VAR_INPUT
  IN0 : INT ;
  IN1 : WORD ;
  IN2 : INT ;
  IN3 : INT ;
END_VAR
VAR_OUTPUT
  OUT4 : BOOL ;
  OUT5 : WORD ;
END_VAR
VAR
  STAT6 : STRUCT
   STAT7 : WORD ;
   STAT8 : WORD ;
   STAT9 : WORD ;
   STAT10 : BYTE ;
   STAT11 : BYTE ;
   STAT12 : BYTE ;
   STAT13 : BYTE ;
   STAT14 : BYTE ;
   STAT15 : BYTE ;
   STAT16 : BYTE ;
   STAT17 : BYTE ;
   STAT18 : BYTE ;
   STAT19 : BYTE ;
   STAT20 : BYTE ;
   STAT21 : BYTE ;
   STAT22 : BYTE ;
   STAT23 : BYTE ;
   STAT24 : BYTE ;
   STAT25 : BYTE ;
   STAT26 : BYTE ;
   STAT27 : BYTE ;
   STAT28 : BYTE ;
   STAT29 : BYTE ;
   STAT30 : BYTE ;
   STAT31 : BYTE ;
   STAT32 : BYTE ;
   STAT33 : BYTE ;
   STAT34 : BYTE ;
   STAT35 : BYTE ;
   STAT36 : BYTE ;
   STAT37 : BYTE ;
   STAT38 : BYTE ;
   STAT39 : BYTE ;
   STAT40 : BYTE ;
   STAT41 : BYTE ;
   STAT42 : BYTE ;
   STAT43 : BYTE ;
   STAT44 : BYTE ;
   STAT45 : BYTE ;
   STAT46 : BYTE ;
   STAT47 : BYTE ;
   STAT48 : BYTE ;
   STAT49 : BYTE ;
   STAT50 : BYTE ;
   STAT51 : BYTE ;
   STAT52 : BYTE ;
   STAT53 : BYTE ;
   STAT54 : BYTE ;
   STAT55 : BYTE ;
   STAT56 : BYTE ;
   STAT57 : BYTE ;
   STAT58 : BYTE ;
   STAT59 : BYTE ;
   STAT60 : BYTE ;
   STAT61 : BYTE ;
   STAT62 : BYTE ;
   STAT63 : BYTE ;
   STAT64 : BYTE ;
   STAT65 : BYTE ;
   STAT66 : BYTE ;
   STAT67 : BYTE ;
   STAT68 : BYTE ;
   STAT69 : BYTE ;
   STAT70 : BYTE ;
   STAT71 : BYTE ;
   STAT72 : BYTE ;
   STAT73 : BYTE ;
   STAT74 : BYTE ;
   STAT75 : BYTE ;
   STAT76 : BYTE ;
   STAT77 : BYTE ;
   STAT78 : BYTE ;
   STAT79 : BYTE ;
   STAT80 : BYTE ;
   STAT81 : BYTE ;
   STAT82 : BYTE ;
   STAT83 : BYTE ;
   STAT84 : BYTE ;
   STAT85 : BYTE ;
   STAT86 : BYTE ;
   STAT87 : BYTE ;
   STAT88 : BYTE ;
   STAT89 : BYTE ;
   STAT90 : BYTE ;
   STAT91 : BYTE ;
   STAT92 : BYTE ;
   STAT93 : BYTE ;
   STAT94 : BYTE ;
   STAT95 : BYTE ;
   STAT96 : BYTE ;
   STAT97 : BYTE ;
   STAT98 : BYTE ;
   STAT99 : BYTE ;
   STAT100 : BYTE ;
   STAT101 : BYTE ;
   STAT102 : BYTE ;
   STAT103 : BYTE ;
   STAT104 : BYTE ;
   STAT105 : BYTE ;
   STAT106 : BYTE ;
   STAT107 : BYTE ;
   STAT108 : BYTE ;
   STAT109 : BYTE ;
   STAT110 : BYTE ;
   STAT111 : BYTE ;
   STAT112 : BYTE ;
   STAT113 : BYTE ;
   STAT114 : BYTE ;
   STAT115 : BYTE ;
   STAT116 : BYTE ;
   STAT117 : BYTE ;
   STAT118 : BYTE ;
   STAT119 : BYTE ;
   STAT120 : BYTE ;
   STAT121 : BYTE ;
   STAT122 : BYTE ;
   STAT123 : BYTE ;
   STAT124 : BYTE ;
   STAT125 : BYTE ;
   STAT126 : BYTE ;
   STAT127 : BYTE ;
   STAT128 : BYTE ;
   STAT129 : BYTE ;
   STAT130 : BYTE ;
   STAT131 : BYTE ;
   STAT132 : BYTE ;
   STAT133 : BYTE ;
   STAT134 : BYTE ;
   STAT135 : BYTE ;
   STAT136 : BYTE ;
   STAT137 : BYTE ;
   STAT138 : BYTE ;
   STAT139 : BYTE ;
   STAT140 : BYTE ;
   STAT141 : BYTE ;
   STAT142 : BYTE ;
   STAT143 : BYTE ;
   STAT144 : BYTE ;
   STAT145 : BYTE ;
   STAT146 : BYTE ;
   STAT147 : BYTE ;
   STAT148 : BYTE ;
   STAT149 : BYTE ;
   STAT150 : BYTE ;
   STAT151 : BYTE ;
   STAT152 : BYTE ;
   STAT153 : BYTE ;
   STAT154 : BYTE ;
   STAT155 : BYTE ;
   STAT156 : BYTE ;
   STAT157 : BYTE ;
   STAT158 : BYTE ;
   STAT159 : BYTE ;
   STAT160 : BYTE ;
   STAT161 : BYTE ;
   STAT162 : BYTE ;
   STAT163 : BYTE ;
   STAT164 : BYTE ;
   STAT165 : BYTE ;
   STAT166 : BYTE ;
   STAT167 : BYTE ;
   STAT168 : BYTE ;
   STAT169 : BYTE ;
   STAT170 : BYTE ;
   STAT171 : BYTE ;
   STAT172 : BYTE ;
   STAT173 : BYTE ;
   STAT174 : BYTE ;
   STAT175 : BYTE ;
   STAT176 : BYTE ;
   STAT177 : BYTE ;
   STAT178 : BYTE ;
   STAT179 : BYTE ;
   STAT180 : BYTE ;
   STAT181 : BYTE ;
   STAT182 : BYTE ;
   STAT183 : BYTE ;
   STAT184 : BYTE ;
   STAT185 : BYTE ;
   STAT186 : BYTE ;
   STAT187 : BYTE ;
   STAT188 : BYTE ;
   STAT189 : BYTE ;
   STAT190 : BYTE ;
   STAT191 : BYTE ;
   STAT192 : BYTE ;
   STAT193 : BYTE ;
   STAT194 : BYTE ;
   STAT195 : BYTE ;
   STAT196 : BYTE ;
   STAT197 : BYTE ;
   STAT198 : BYTE ;
   STAT199 : BYTE ;
   STAT200 : BYTE ;
   STAT201 : BYTE ;
   STAT202 : BYTE ;
   STAT203 : BYTE ;
   STAT204 : BYTE ;
   STAT205 : BYTE ;
   STAT206 : BYTE ;
   STAT207 : BYTE ;
   STAT208 : BYTE ;
   STAT209 : BYTE ;
   STAT210 : BYTE ;
   STAT211 : BYTE ;
   STAT212 : BYTE ;
   STAT213 : BYTE ;
   STAT214 : BYTE ;
   STAT215 : BYTE ;
   STAT216 : BYTE ;
   STAT217 : BYTE ;
   STAT218 : BYTE ;
   STAT219 : BYTE ;
   STAT220 : BYTE ;
   STAT221 : BYTE ;
   STAT222 : BYTE ;
   STAT223 : BYTE ;
   STAT224 : BYTE ;
   STAT225 : BYTE ;
   STAT226 : BYTE ;
   STAT227 : BYTE ;
   STAT228 : BYTE ;
   STAT229 : BYTE ;
   STAT230 : BYTE ;
   STAT231 : BYTE ;
   STAT232 : BYTE ;
   STAT233 : BYTE ;
   STAT234 : BYTE ;
   STAT235 : BYTE ;
   STAT236 : BYTE ;
   STAT237 : BYTE ;
   STAT238 : BYTE ;
   STAT239 : BYTE ;
   STAT240 : BYTE ;
   STAT241 : BYTE ;
   STAT242 : BYTE ;
   STAT243 : BYTE ;
   STAT244 : BYTE ;
   STAT245 : BYTE ;
   STAT246 : BYTE ;
   STAT247 : BYTE ;
   STAT248 : BYTE ;
   STAT249 : BYTE ;
   STAT250 : BYTE ;
   STAT251 : BYTE ;
   STAT252 : BYTE ;
   STAT253 : BYTE ;
   STAT254 : BYTE ;
   STAT255 : BYTE ;
   STAT256 : BYTE ;
   STAT257 : BYTE ;
   STAT258 : BYTE ;
   STAT259 : BYTE ;
   STAT260 : BYTE ;
  END_STRUCT ;
  STAT261 : STRUCT
   STAT262 : WORD ;
   STAT263 : WORD ;
   STAT264 : WORD ;
   STAT265 : BYTE ;
   STAT266 : BYTE ;
   STAT267 : WORD ;
   STAT268 : WORD ;
   STAT269 : BYTE ;
   STAT270 : BYTE ;
   STAT271 : BYTE ;
   STAT272 : BYTE ;
   STAT273 : BYTE ;
   STAT274 : BYTE ;
   STAT275 : BYTE ;
   STAT276 : BYTE ;
   STAT277 : BYTE ;
   STAT278 : BYTE ;
   STAT279 : BYTE ;
   STAT280 : BYTE ;
   STAT281 : BYTE ;
   STAT282 : BYTE ;
   STAT283 : BYTE ;
   STAT284 : BYTE ;
   STAT285 : BYTE ;
   STAT286 : BYTE ;
   STAT287 : BYTE ;
   STAT288 : BYTE ;
   STAT289 : BYTE ;
   STAT290 : BYTE ;
   STAT291 : BYTE ;
   STAT292 : BYTE ;
   STAT293 : BYTE ;
   STAT294 : BYTE ;
   STAT295 : BYTE ;
   STAT296 : BYTE ;
   STAT297 : BYTE ;
   STAT298 : BYTE ;
   STAT299 : BYTE ;
   STAT300 : BYTE ;
   STAT301 : BYTE ;
   STAT302 : BYTE ;
   STAT303 : BYTE ;
   STAT304 : BYTE ;
   STAT305 : BYTE ;
   STAT306 : BYTE ;
   STAT307 : BYTE ;
   STAT308 : BYTE ;
   STAT309 : BYTE ;
   STAT310 : BYTE ;
   STAT311 : BYTE ;
   STAT312 : BYTE ;
   STAT313 : BYTE ;
   STAT314 : BYTE ;
   STAT315 : BYTE ;
   STAT316 : BYTE ;
   STAT317 : BYTE ;
   STAT318 : BYTE ;
   STAT319 : BYTE ;
   STAT320 : BYTE ;
   STAT321 : BYTE ;
   STAT322 : BYTE ;
   STAT323 : BYTE ;
   STAT324 : BYTE ;
   STAT325 : BYTE ;
   STAT326 : BYTE ;
   STAT327 : BYTE ;
   STAT328 : BYTE ;
   STAT329 : BYTE ;
   STAT330 : BYTE ;
   STAT331 : BYTE ;
   STAT332 : BYTE ;
   STAT333 : BYTE ;
   STAT334 : BYTE ;
   STAT335 : BYTE ;
   STAT336 : BYTE ;
   STAT337 : BYTE ;
   STAT338 : BYTE ;
   STAT339 : BYTE ;
   STAT340 : BYTE ;
   STAT341 : BYTE ;
   STAT342 : BYTE ;
   STAT343 : BYTE ;
   STAT344 : BYTE ;
   STAT345 : BYTE ;
   STAT346 : BYTE ;
   STAT347 : BYTE ;
   STAT348 : BYTE ;
   STAT349 : BYTE ;
   STAT350 : BYTE ;
   STAT351 : BYTE ;
   STAT352 : BYTE ;
   STAT353 : BYTE ;
   STAT354 : BYTE ;
   STAT355 : BYTE ;
   STAT356 : BYTE ;
   STAT357 : BYTE ;
   STAT358 : BYTE ;
   STAT359 : BYTE ;
   STAT360 : BYTE ;
   STAT361 : BYTE ;
   STAT362 : BYTE ;
   STAT363 : BYTE ;
   STAT364 : BYTE ;
   STAT365 : BYTE ;
   STAT366 : BYTE ;
   STAT367 : BYTE ;
   STAT368 : BYTE ;
   STAT369 : BYTE ;
   STAT370 : BYTE ;
   STAT371 : BYTE ;
   STAT372 : BYTE ;
   STAT373 : BYTE ;
   STAT374 : BYTE ;
   STAT375 : BYTE ;
   STAT376 : BYTE ;
   STAT377 : BYTE ;
   STAT378 : BYTE ;
   STAT379 : BYTE ;
   STAT380 : BYTE ;
   STAT381 : BYTE ;
   STAT382 : BYTE ;
   STAT383 : BYTE ;
   STAT384 : BYTE ;
   STAT385 : BYTE ;
   STAT386 : BYTE ;
   STAT387 : BYTE ;
   STAT388 : BYTE ;
   STAT389 : BYTE ;
   STAT390 : BYTE ;
   STAT391 : BYTE ;
   STAT392 : BYTE ;
   STAT393 : BYTE ;
   STAT394 : BYTE ;
   STAT395 : BYTE ;
   STAT396 : BYTE ;
   STAT397 : BYTE ;
   STAT398 : BYTE ;
   STAT399 : BYTE ;
   STAT400 : BYTE ;
   STAT401 : BYTE ;
   STAT402 : BYTE ;
   STAT403 : BYTE ;
   STAT404 : BYTE ;
   STAT405 : BYTE ;
   STAT406 : BYTE ;
   STAT407 : BYTE ;
   STAT408 : BYTE ;
   STAT409 : BYTE ;
   STAT410 : BYTE ;
   STAT411 : BYTE ;
   STAT412 : BYTE ;
   STAT413 : BYTE ;
   STAT414 : BYTE ;
   STAT415 : BYTE ;
   STAT416 : BYTE ;
   STAT417 : BYTE ;
   STAT418 : BYTE ;
   STAT419 : BYTE ;
   STAT420 : BYTE ;
   STAT421 : BYTE ;
   STAT422 : BYTE ;
   STAT423 : BYTE ;
   STAT424 : BYTE ;
   STAT425 : BYTE ;
   STAT426 : BYTE ;
   STAT427 : BYTE ;
   STAT428 : BYTE ;
   STAT429 : BYTE ;
   STAT430 : BYTE ;
   STAT431 : BYTE ;
   STAT432 : BYTE ;
   STAT433 : BYTE ;
   STAT434 : BYTE ;
   STAT435 : BYTE ;
   STAT436 : BYTE ;
   STAT437 : BYTE ;
   STAT438 : BYTE ;
   STAT439 : BYTE ;
   STAT440 : BYTE ;
   STAT441 : BYTE ;
   STAT442 : BYTE ;
   STAT443 : BYTE ;
   STAT444 : BYTE ;
   STAT445 : BYTE ;
   STAT446 : BYTE ;
   STAT447 : BYTE ;
   STAT448 : BYTE ;
   STAT449 : BYTE ;
   STAT450 : BYTE ;
   STAT451 : BYTE ;
   STAT452 : BYTE ;
   STAT453 : BYTE ;
   STAT454 : BYTE ;
   STAT455 : BYTE ;
   STAT456 : BYTE ;
   STAT457 : BYTE ;
   STAT458 : BYTE ;
   STAT459 : BYTE ;
   STAT460 : BYTE ;
   STAT461 : BYTE ;
   STAT462 : BYTE ;
   STAT463 : BYTE ;
   STAT464 : BYTE ;
   STAT465 : BYTE ;
   STAT466 : BYTE ;
   STAT467 : BYTE ;
   STAT468 : BYTE ;
   STAT469 : BYTE ;
   STAT470 : BYTE ;
   STAT471 : BYTE ;
   STAT472 : BYTE ;
   STAT473 : BYTE ;
   STAT474 : BYTE ;
   STAT475 : BYTE ;
   STAT476 : BYTE ;
   STAT477 : BYTE ;
   STAT478 : BYTE ;
   STAT479 : BYTE ;
   STAT480 : BYTE ;
   STAT481 : BYTE ;
   STAT482 : BYTE ;
   STAT483 : BYTE ;
   STAT484 : BYTE ;
   STAT485 : BYTE ;
   STAT486 : BYTE ;
   STAT487 : BYTE ;
   STAT488 : BYTE ;
   STAT489 : BYTE ;
   STAT490 : BYTE ;
   STAT491 : BYTE ;
   STAT492 : BYTE ;
   STAT493 : BYTE ;
   STAT494 : BYTE ;
   STAT495 : BYTE ;
   STAT496 : BYTE ;
   STAT497 : BYTE ;
   STAT498 : BYTE ;
   STAT499 : BYTE ;
   STAT500 : BYTE ;
   STAT501 : BYTE ;
   STAT502 : BYTE ;
   STAT503 : BYTE ;
   STAT504 : BYTE ;
   STAT505 : BYTE ;
   STAT506 : BYTE ;
   STAT507 : BYTE ;
   STAT508 : BYTE ;
   STAT509 : BYTE ;
   STAT510 : BYTE ;
   STAT511 : BYTE ;
   STAT512 : BYTE ;
   STAT513 : BYTE ;
   STAT514 : BYTE ;
  END_STRUCT ;
  STAT515 : INT ;
  STAT516 : INT ;
  STAT517 : BOOL ;
  STAT518 : BOOL ;
  STAT519 : BOOL ;
  STAT520 : BOOL ;
  STAT521 : WORD ;
  STAT522 : INT ;
  STAT523 : BOOL ;
  STAT524 : BOOL ;
  STAT525 : WORD ;
  STAT526 : INT ;
  STAT527 : INT ;
  STAT528 : BOOL ;
  STAT529 : BOOL ;
  STAT530 : WORD ;
  STAT531 : BOOL ;
  STAT532 : WORD ;
  STAT533 : "TON";
  STAT541 : BOOL ;
  STAT542 : BOOL ;
  STAT543 : BOOL ;
  STAT544 : WORD ;
END_VAR
VAR_TEMP
  TEMP545 : ANY ;
  TEMP546 : ANY ;
  TEMP547 : INT ;
  TEMP548 : DWORD ;
  TEMP549 : DWORD ;
END_VAR
BEGIN
NETWORK
TITLE =
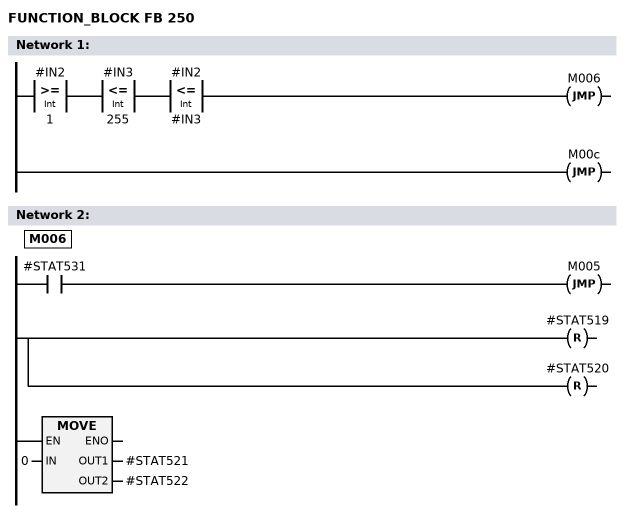

      SET   ;
      A(    ;
      L     #IN2;
      L     1;
      >=I   ;
      )     ;
      A(    ;
      L     #IN3;
      L     255;
      <=I   ;
      )     ;
      A(    ;
      L     #IN2;
      L     #IN3;
      <=I   ;
      )     ;
      JC    M006;
      JU    M00c;
NETWORK
TITLE =

M006: A     #STAT531;
      JC    M005;
      SET   ;
      R     #STAT519;
      R     #STAT520;
      L     0;
      T     #STAT521;
      T     #STAT522;
NETWORK
TITLE =

      LAR1  P##TEMP545;
      L     B#16#10;
      T     LB [AR1,P#0.0];
      L     B#16#2;
      T     LB [AR1,P#1.0];
      L     6;
      T     LW [AR1,P#2.0];
      L     DINO;
      T     LW [AR1,P#4.0];
      L     270;
      L     8;
      *I    ;
      L     P#DBX 0.0;
      +D    ;
      T     LD [AR1,P#6.0];
NETWORK
TITLE =
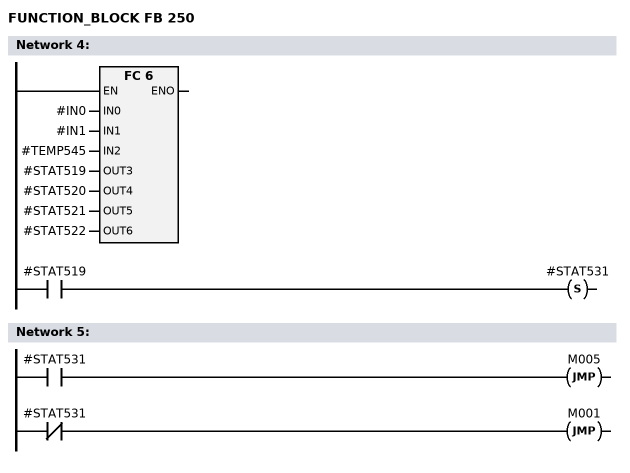

      CALL FC     6 (
           IN0                      := #IN0,
           IN1                      := #IN1,
           IN2                      := #TEMP545,
           OUT3                     := #STAT519,
           OUT4                     := #STAT520,
           OUT5                     := #STAT521,
           OUT6                     := #STAT522);
      SET   ;
      A     #STAT519;
      S     #STAT531;
NETWORK
TITLE =

      A     #STAT531;
      JC    M005;
      AN    #STAT531;
      JC    M001;
NETWORK
TITLE =

M005: LAR1  P##TEMP546;
      L     B#16#10;
      T     LB [AR1,P#0.0];
      L     B#16#2;
      T     LB [AR1,P#1.0];
      L     DIW  274;
      T     LW [AR1,P#2.0];
      L     DINO;
      T     LW [AR1,P#4.0];
      L     276;
      L     8;
      *I    ;
      L     P#DBX 0.0;
      +D    ;
      T     LD [AR1,P#6.0];
NETWORK
TITLE =
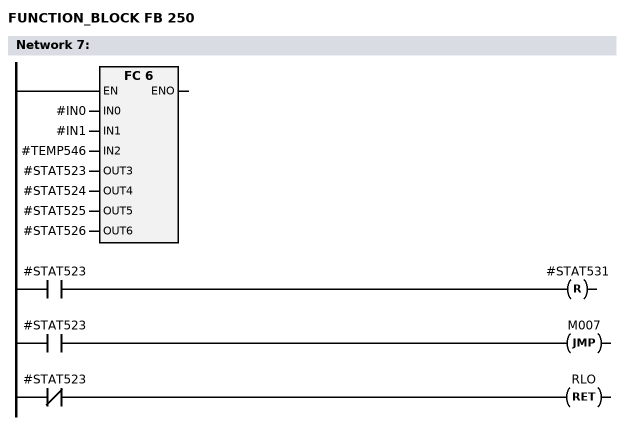

      CALL FC     6 (
           IN0                      := #IN0,
           IN1                      := #IN1,
           IN2                      := #TEMP546,
           OUT3                     := #STAT523,
           OUT4                     := #STAT524,
           OUT5                     := #STAT525,
           OUT6                     := #STAT526);
      SET   ;
      A     #STAT523;
      R     #STAT531;
      A     #STAT523;
      JC    M007;
      AN    #STAT523;
      BEC   ;
NETWORK
TITLE =

M007: SET   ;
      L     #STAT261.STAT266;
      L     3;
      ==I   ;
      =     #STAT517;
      L     #STAT261.STAT266;
      L     16;
      ==I   ;
      =     #STAT518;
      A     #STAT517;
      JC    M00b;
      A     #STAT518;
      JC    M009;
      JU    M008;
NETWORK
TITLE =

M00b: O(    ;
      L     #STAT261.STAT268;
      L     1;
      <I    ;
      )     ;
      O(    ;
      L     #STAT261.STAT268;
      L     100;
      >I    ;
      )     ;
      JC    M00a;
      L     #STAT261.STAT267;
      SRW   8;
      T     #TEMP547;
      L     #IN2;
      L     #TEMP547;
      +I    ;
      T     #TEMP547;
      O(    ;
      L     #TEMP547;
      L     #IN2;
      <I    ;
      )     ;
      O(    ;
      L     #TEMP547;
      L     #IN3;
      >I    ;
      )     ;
      JC    M00a;
      L     #STAT261.STAT262;
      T     #STAT6.STAT7;
      L     #STAT261.STAT263;
      T     #STAT6.STAT8;
      L     #STAT261.STAT265;
      T     #STAT6.STAT10;
      L     #STAT261.STAT266;
      T     #STAT6.STAT11;
      L     #STAT261.STAT268;
      SLW   1;
      T     #STAT6.STAT12;
      L     #STAT6.STAT12;
      +     3;
      T     #STAT6.STAT9;
      OPN   DB [#TEMP547];
      L     #STAT261.STAT267;
      SLW   8;
      SRW   8;
      SLD   4;
      T     #TEMP548;
      L     P##STAT6;
      L     P#9.0;
      +D    ;
      T     #TEMP549;
      L     #STAT261.STAT268;
M003: T     #STAT532;
      L     DBW [#TEMP548];
      T     DIW [#TEMP549];
      L     #TEMP548;
      +     16;
      T     #TEMP548;
      L     #TEMP549;
      +     16;
      T     #TEMP549;
      L     #STAT532;
      LOOP  M003;
      L     #STAT6.STAT9;
      +     6;
      T     #STAT527;
      L     W#16#0;
      T     #OUT5;
      R     #OUT4;
      S     #STAT543;
      JU    M001;
NETWORK
TITLE =

M009: O(    ;
      L     #STAT261.STAT268;
      L     1;
      <I    ;
      )     ;
      O(    ;
      L     #STAT261.STAT268;
      L     100;
      >I    ;
      )     ;
      JC    M00a;
      L     #STAT261.STAT267;
      T     #STAT6.STAT15;
      SRW   8;
      T     #STAT6.STAT12;
      T     #TEMP547;
      L     #IN2;
      L     #TEMP547;
      +I    ;
      T     #TEMP547;
      O(    ;
      L     #TEMP547;
      L     #IN2;
      <I    ;
      )     ;
      O(    ;
      L     #TEMP547;
      L     #IN3;
      >I    ;
      )     ;
      JC    M00a;
      L     #STAT261.STAT262;
      T     #STAT6.STAT7;
      L     #STAT261.STAT263;
      T     #STAT6.STAT8;
      L     #STAT261.STAT265;
      T     #STAT6.STAT10;
      L     #STAT261.STAT266;
      T     #STAT6.STAT11;
      L     6;
      T     #STAT6.STAT9;
      L     0;
      T     #STAT6.STAT14;
      L     #STAT261.STAT268;
      T     #STAT6.STAT15;
      OPN   DB [#TEMP547];
      L     #STAT261.STAT267;
      SLW   8;
      SRW   8;
      T     #STAT6.STAT13;
      SLD   4;
      T     #TEMP549;
      L     P##STAT261;
      L     P#13.0;
      +D    ;
      T     #TEMP548;
      L     #STAT261.STAT268;
M004: T     #STAT532;
      L     DIW [#TEMP548];
      T     DBW [#TEMP549];
      L     #TEMP548;
      +     16;
      T     #TEMP548;
      L     #TEMP549;
      +     16;
      T     #TEMP549;
      L     #STAT532;
      LOOP  M004;
      L     12;
      T     #STAT527;
      L     W#16#0;
      T     #OUT5;
      R     #OUT4;
      S     #STAT543;
      JU    M001;
NETWORK
TITLE =

M00c: L     W#16#290;
      T     #OUT5;
      S     #OUT4;
      BEU   ;
M008: L     B#16#1;
      T     #STAT6.STAT12;
      L     W#16#300;
      T     #OUT5;
      JU    M002;
M00a: L     B#16#2;
      T     #STAT6.STAT12;
      L     W#16#381;
      T     #OUT5;
      JU    M002;
M002: L     #STAT261.STAT262;
      T     #STAT6.STAT7;
      L     #STAT261.STAT263;
      T     #STAT6.STAT8;
      L     #STAT261.STAT265;
      T     #STAT6.STAT10;
      L     #STAT261.STAT266;
      +     B#16#80;
      T     #STAT6.STAT11;
      L     3;
      T     #STAT6.STAT9;
      L     9;
      T     #STAT527;
      S     #OUT4;
      S     #STAT543;
      JU    M001;
NETWORK
TITLE =

M001: CALL FC     5 (
           IN0                      := #STAT543,
           IN1                      := #IN0,
           IN2                      := #IN1,
           IN3                      := #STAT6,
           IN4                      := #STAT527,
           OUT5                     := #STAT528,
           OUT6                     := #STAT529,
           OUT7                     := #STAT530);
      SET   ;
      R     #STAT543;
      BEU   ;
END_FUNCTION_BLOCK

FUNCTION FC 14 : VOID
VERSION : 0.1

BEGIN
NETWORK
TITLE =

      CALL FB   250 , DB   250 (
           IN0                      := 1,
           IN1                      := W#16#180,
           IN2                      := 95,
           IN3                      := 95,
           OUT4                     := DB250.DBX    8.0,
           OUT5                     := DB250.DBW   10);
      NOP   0;
NETWORK
TITLE =

      A     I      0.0;
      =     DB95.DBX    1.0;
NETWORK
TITLE =

      A     Q    160.6;
      =     DB95.DBX    1.1;
NETWORK
TITLE =

      A(    ;
      L     DB51.DBD  252;
      L     1.000000e+003;
      *R    ;
      T     MD   100;
      AN    OV;
      SAVE  ;
      CLR   ;
      A     BR;
      )     ;
      JNB   M001;
      L     MD   100;
      RND   ;
      T     DB95.DBW   18;
M001: NOP   0;
NETWORK
TITLE =

      A(    ;
      L     DB51.DBD  292;
      L     1.000000e+003;
      *R    ;
      T     MD   104;
      AN    OV;
      SAVE  ;
      CLR   ;
      A     BR;
      )     ;
      JNB   M002;
      L     MD   104;
      RND   ;
      T     DB95.DBW   20;
M002: NOP   0;
NETWORK
TITLE =

      A(    ;
      L     DB51.DBD   92;
      L     1.000000e+003;
      *R    ;
      T     MD   108;
      AN    OV;
      SAVE  ;
      CLR   ;
      A     BR;
      )     ;
      JNB   M003;
      L     MD   108;
      RND   ;
      T     DB95.DBW   22;
M003: NOP   0;
NETWORK
TITLE =

      A(    ;
      L     DB51.DBD  212;
      L     1.000000e+003;
      *R    ;
      T     MD   112;
      AN    OV;
      SAVE  ;
      CLR   ;
      A     BR;
      )     ;
      JNB   M004;
      L     MD   112;
      RND   ;
      T     DB95.DBW   24;
M004: NOP   0;
NETWORK
TITLE =

      A(    ;
      L     DB51.DBD   52;
      L     1.000000e+003;
      *R    ;
      T     MD   116;
      AN    OV;
      SAVE  ;
      CLR   ;
      A     BR;
      )     ;
      JNB   M005;
      L     MD   116;
      RND   ;
      T     DB95.DBW   26;
M005: NOP   0;
NETWORK
TITLE =

      A(    ;
      L     DB51.DBD  172;
      L     1.000000e+003;
      *R    ;
      T     MD   120;
      AN    OV;
      SAVE  ;
      CLR   ;
      A     BR;
      )     ;
      JNB   M006;
      L     MD   120;
      RND   ;
      T     DB95.DBW   28;
M006: NOP   0;
NETWORK
TITLE =

      A(    ;
      L     DB51.DBD   12;
      L     1.000000e+003;
      *R    ;
      T     MD   124;
      AN    OV;
      SAVE  ;
      CLR   ;
      A     BR;
      )     ;
      JNB   M007;
      L     MD   124;
      RND   ;
      T     DB95.DBW   30;
M007: NOP   0;
NETWORK
TITLE =

      A(    ;
      L     DB51.DBD  132;
      L     1.000000e+003;
      *R    ;
      T     MD   128;
      AN    OV;
      SAVE  ;
      CLR   ;
      A     BR;
      )     ;
      JNB   M008;
      L     MD   128;
      RND   ;
      T     DB95.DBW   32;
M008: NOP   0;
NETWORK
TITLE =

      A(    ;
      L     DB51.DBD  256;
      L     1.000000e+003;
      *R    ;
      T     MD   132;
      AN    OV;
      SAVE  ;
      CLR   ;
      A     BR;
      )     ;
      JNB   M009;
      L     MD   132;
      RND   ;
      T     DB95.DBW   38;
M009: NOP   0;
NETWORK
TITLE =

      A(    ;
      L     DB51.DBD  296;
      L     1.000000e+003;
      *R    ;
      T     MD   136;
      AN    OV;
      SAVE  ;
      CLR   ;
      A     BR;
      )     ;
      JNB   M00a;
      L     MD   136;
      RND   ;
      T     DB95.DBW   40;
M00a: NOP   0;
NETWORK
TITLE =

      A(    ;
      L     DB51.DBD   96;
      L     1.000000e+003;
      *R    ;
      T     MD   140;
      AN    OV;
      SAVE  ;
      CLR   ;
      A     BR;
      )     ;
      JNB   M00b;
      L     MD   140;
      RND   ;
      T     DB95.DBW   42;
M00b: NOP   0;
NETWORK
TITLE =

      A(    ;
      L     DB51.DBD  216;
      L     1.000000e+003;
      *R    ;
      T     MD   144;
      AN    OV;
      SAVE  ;
      CLR   ;
      A     BR;
      )     ;
      JNB   M00c;
      L     MD   144;
      RND   ;
      T     DB95.DBW   44;
M00c: NOP   0;
NETWORK
TITLE =

      A(    ;
      L     DB51.DBD   56;
      L     1.000000e+003;
      *R    ;
      T     MD   148;
      AN    OV;
      SAVE  ;
      CLR   ;
      A     BR;
      )     ;
      JNB   M00d;
      L     MD   148;
      RND   ;
      T     DB95.DBW   46;
M00d: NOP   0;
NETWORK
TITLE =

      A(    ;
      L     DB51.DBD  176;
      L     1.000000e+003;
      *R    ;
      T     MD   152;
      AN    OV;
      SAVE  ;
      CLR   ;
      A     BR;
      )     ;
      JNB   M00e;
      L     MD   152;
      RND   ;
      T     DB95.DBW   48;
M00e: NOP   0;
NETWORK
TITLE =

      A(    ;
      L     DB51.DBD   16;
      L     1.000000e+003;
      *R    ;
      T     MD   156;
      AN    OV;
      SAVE  ;
      CLR   ;
      A     BR;
      )     ;
      JNB   M00f;
      L     MD   156;
      RND   ;
      T     DB95.DBW   50;
M00f: NOP   0;
NETWORK
TITLE =

      A(    ;
      L     DB51.DBD  136;
      L     1.000000e+003;
      *R    ;
      T     MD   160;
      AN    OV;
      SAVE  ;
      CLR   ;
      A     BR;
      )     ;
      JNB   M010;
      L     MD   160;
      RND   ;
      T     DB95.DBW   52;
M010: NOP   0;
NETWORK
TITLE =

      A(    ;
      L     DB51.DBD  260;
      L     1.000000e+003;
      *R    ;
      T     MD   164;
      AN    OV;
      SAVE  ;
      CLR   ;
      A     BR;
      )     ;
      JNB   M011;
      L     MD   164;
      RND   ;
      T     DB95.DBW   58;
M011: NOP   0;
NETWORK
TITLE =

      A(    ;
      L     DB51.DBD  300;
      L     1.000000e+003;
      *R    ;
      T     MD   168;
      AN    OV;
      SAVE  ;
      CLR   ;
      A     BR;
      )     ;
      JNB   M012;
      L     MD   168;
      RND   ;
      T     DB95.DBW   60;
M012: NOP   0;
NETWORK
TITLE =

      A(    ;
      L     DB51.DBD  100;
      L     1.000000e+003;
      *R    ;
      T     MD   172;
      AN    OV;
      SAVE  ;
      CLR   ;
      A     BR;
      )     ;
      JNB   M013;
      L     MD   172;
      RND   ;
      T     DB95.DBW   62;
M013: NOP   0;
NETWORK
TITLE =

      A(    ;
      L     DB51.DBD  220;
      L     1.000000e+003;
      *R    ;
      T     MD   176;
      AN    OV;
      SAVE  ;
      CLR   ;
      A     BR;
      )     ;
      JNB   M014;
      L     MD   176;
      RND   ;
      T     DB95.DBW   64;
M014: NOP   0;
NETWORK
TITLE =

      A(    ;
      L     DB51.DBD   60;
      L     1.000000e+003;
      *R    ;
      T     MD   180;
      AN    OV;
      SAVE  ;
      CLR   ;
      A     BR;
      )     ;
      JNB   M015;
      L     MD   180;
      RND   ;
      T     DB95.DBW   66;
M015: NOP   0;
NETWORK
TITLE =

      A(    ;
      L     DB51.DBD  180;
      L     1.000000e+003;
      *R    ;
      T     MD   184;
      AN    OV;
      SAVE  ;
      CLR   ;
      A     BR;
      )     ;
      JNB   M016;
      L     MD   184;
      RND   ;
      T     DB95.DBW   68;
M016: NOP   0;
NETWORK
TITLE =

      A(    ;
      L     DB51.DBD   20;
      L     1.000000e+003;
      *R    ;
      T     MD   188;
      AN    OV;
      SAVE  ;
      CLR   ;
      A     BR;
      )     ;
      JNB   M017;
      L     MD   188;
      RND   ;
      T     DB95.DBW   70;
M017: NOP   0;
NETWORK
TITLE =

      A(    ;
      L     DB51.DBD  140;
      L     1.000000e+003;
      *R    ;
      T     MD   192;
      AN    OV;
      SAVE  ;
      CLR   ;
      A     BR;
      )     ;
      JNB   M018;
      L     MD   192;
      RND   ;
      T     DB95.DBW   72;
M018: NOP   0;
NETWORK
TITLE =

      A(    ;
      L     DB51.DBD  264;
      L     1.000000e+003;
      *R    ;
      T     MD   296;
      AN    OV;
      SAVE  ;
      CLR   ;
      A     BR;
      )     ;
      JNB   M019;
      L     MD   296;
      RND   ;
      T     DB95.DBW   78;
M019: NOP   0;
NETWORK
TITLE =

      A(    ;
      L     DB51.DBD  304;
      L     1.000000e+003;
      *R    ;
      T     MD   304;
      AN    OV;
      SAVE  ;
      CLR   ;
      A     BR;
      )     ;
      JNB   M01a;
      L     MD   304;
      RND   ;
      T     DB95.DBW   80;
M01a: NOP   0;
NETWORK
TITLE =

      A(    ;
      L     DB51.DBD  104;
      L     1.000000e+003;
      *R    ;
      T     MD   308;
      AN    OV;
      SAVE  ;
      CLR   ;
      A     BR;
      )     ;
      JNB   M01b;
      L     MD   308;
      RND   ;
      T     DB95.DBW   82;
M01b: NOP   0;
NETWORK
TITLE =

      A(    ;
      L     DB51.DBD  224;
      L     1.000000e+003;
      *R    ;
      T     MD   312;
      AN    OV;
      SAVE  ;
      CLR   ;
      A     BR;
      )     ;
      JNB   M01c;
      L     MD   312;
      RND   ;
      T     DB95.DBW   84;
M01c: NOP   0;
NETWORK
TITLE =

      A(    ;
      L     DB51.DBD   64;
      L     1.000000e+003;
      *R    ;
      T     MD   316;
      AN    OV;
      SAVE  ;
      CLR   ;
      A     BR;
      )     ;
      JNB   M01d;
      L     MD   316;
      RND   ;
      T     DB95.DBW   86;
M01d: NOP   0;
NETWORK
TITLE =

      A(    ;
      L     DB51.DBD  184;
      L     1.000000e+003;
      *R    ;
      T     MD   320;
      AN    OV;
      SAVE  ;
      CLR   ;
      A     BR;
      )     ;
      JNB   M01e;
      L     MD   320;
      RND   ;
      T     DB95.DBW   88;
M01e: NOP   0;
NETWORK
TITLE =

      A(    ;
      L     DB51.DBD   24;
      L     1.000000e+003;
      *R    ;
      T     MD   324;
      AN    OV;
      SAVE  ;
      CLR   ;
      A     BR;
      )     ;
      JNB   M01f;
      L     MD   324;
      RND   ;
      T     DB95.DBW   90;
M01f: NOP   0;
NETWORK
TITLE =

      A(    ;
      L     DB51.DBD  144;
      L     1.000000e+003;
      *R    ;
      T     MD   328;
      AN    OV;
      SAVE  ;
      CLR   ;
      A     BR;
      )     ;
      JNB   M020;
      L     MD   328;
      RND   ;
      T     DB95.DBW   92;
M020: NOP   0;
END_FUNCTION

FUNCTION FC 1 : VOID
VERSION : 0.1

BEGIN
NETWORK
TITLE =
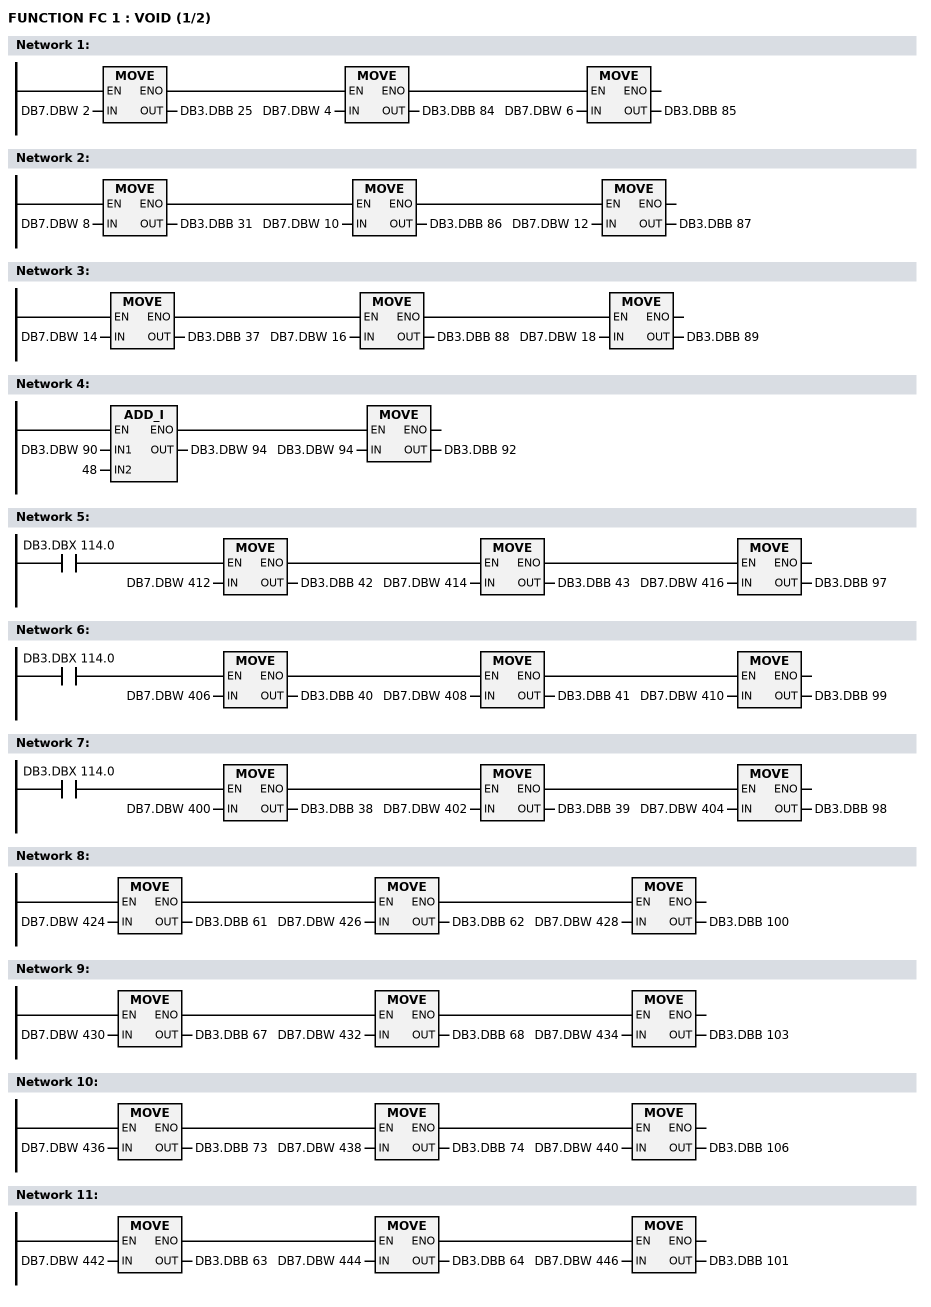

      A(    ;
      A(    ;
      L     DB7.DBW    2;
      T     DB3.DBB   25;
      SET   ;
      SAVE  ;
      CLR   ;
      A     BR;
      )     ;
      JNB   M001;
      L     DB7.DBW    4;
      T     DB3.DBB   84;
      SET   ;
      SAVE  ;
      CLR   ;
M001: A     BR;
      )     ;
      JNB   M002;
      L     DB7.DBW    6;
      T     DB3.DBB   85;
M002: NOP   0;
NETWORK
TITLE =

      A(    ;
      A(    ;
      L     DB7.DBW    8;
      T     DB3.DBB   31;
      SET   ;
      SAVE  ;
      CLR   ;
      A     BR;
      )     ;
      JNB   M003;
      L     DB7.DBW   10;
      T     DB3.DBB   86;
      SET   ;
      SAVE  ;
      CLR   ;
M003: A     BR;
      )     ;
      JNB   M004;
      L     DB7.DBW   12;
      T     DB3.DBB   87;
M004: NOP   0;
NETWORK
TITLE =

      A(    ;
      A(    ;
      L     DB7.DBW   14;
      T     DB3.DBB   37;
      SET   ;
      SAVE  ;
      CLR   ;
      A     BR;
      )     ;
      JNB   M005;
      L     DB7.DBW   16;
      T     DB3.DBB   88;
      SET   ;
      SAVE  ;
      CLR   ;
M005: A     BR;
      )     ;
      JNB   M006;
      L     DB7.DBW   18;
      T     DB3.DBB   89;
M006: NOP   0;
NETWORK
TITLE =

      A(    ;
      L     DB3.DBW   90;
      L     48;
      +I    ;
      T     DB3.DBW   94;
      AN    OV;
      SAVE  ;
      CLR   ;
      A     BR;
      )     ;
      JNB   M007;
      L     DB3.DBW   94;
      T     DB3.DBB   92;
M007: NOP   0;
NETWORK
TITLE =

      A(    ;
      A(    ;
      A     DB3.DBX  114.0;
      JNB   M008;
      L     DB7.DBW  412;
      T     DB3.DBB   42;
      SET   ;
      SAVE  ;
      CLR   ;
M008: A     BR;
      )     ;
      JNB   M009;
      L     DB7.DBW  414;
      T     DB3.DBB   43;
      SET   ;
      SAVE  ;
      CLR   ;
M009: A     BR;
      )     ;
      JNB   M00e;
      L     DB7.DBW  416;
      T     DB3.DBB   97;
M00e: NOP   0;
NETWORK
TITLE =

      A(    ;
      A(    ;
      A     DB3.DBX  114.0;
      JNB   M00f;
      L     DB7.DBW  406;
      T     DB3.DBB   40;
      SET   ;
      SAVE  ;
      CLR   ;
M00f: A     BR;
      )     ;
      JNB   M010;
      L     DB7.DBW  408;
      T     DB3.DBB   41;
      SET   ;
      SAVE  ;
      CLR   ;
M010: A     BR;
      )     ;
      JNB   M011;
      L     DB7.DBW  410;
      T     DB3.DBB   99;
M011: NOP   0;
NETWORK
TITLE =

      A(    ;
      A(    ;
      A     DB3.DBX  114.0;
      JNB   M012;
      L     DB7.DBW  400;
      T     DB3.DBB   38;
      SET   ;
      SAVE  ;
      CLR   ;
M012: A     BR;
      )     ;
      JNB   M013;
      L     DB7.DBW  402;
      T     DB3.DBB   39;
      SET   ;
      SAVE  ;
      CLR   ;
M013: A     BR;
      )     ;
      JNB   M014;
      L     DB7.DBW  404;
      T     DB3.DBB   98;
M014: NOP   0;
NETWORK
TITLE =

      A(    ;
      A(    ;
      L     DB7.DBW  424;
      T     DB3.DBB   61;
      SET   ;
      SAVE  ;
      CLR   ;
      A     BR;
      )     ;
      JNB   M015;
      L     DB7.DBW  426;
      T     DB3.DBB   62;
      SET   ;
      SAVE  ;
      CLR   ;
M015: A     BR;
      )     ;
      JNB   M016;
      L     DB7.DBW  428;
      T     DB3.DBB  100;
M016: NOP   0;
NETWORK
TITLE =

      A(    ;
      A(    ;
      L     DB7.DBW  430;
      T     DB3.DBB   67;
      SET   ;
      SAVE  ;
      CLR   ;
      A     BR;
      )     ;
      JNB   M017;
      L     DB7.DBW  432;
      T     DB3.DBB   68;
      SET   ;
      SAVE  ;
      CLR   ;
M017: A     BR;
      )     ;
      JNB   M018;
      L     DB7.DBW  434;
      T     DB3.DBB  103;
M018: NOP   0;
NETWORK
TITLE =

      A(    ;
      A(    ;
      L     DB7.DBW  436;
      T     DB3.DBB   73;
      SET   ;
      SAVE  ;
      CLR   ;
      A     BR;
      )     ;
      JNB   M019;
      L     DB7.DBW  438;
      T     DB3.DBB   74;
      SET   ;
      SAVE  ;
      CLR   ;
M019: A     BR;
      )     ;
      JNB   M01a;
      L     DB7.DBW  440;
      T     DB3.DBB  106;
M01a: NOP   0;
NETWORK
TITLE =

      A(    ;
      A(    ;
      L     DB7.DBW  442;
      T     DB3.DBB   63;
      SET   ;
      SAVE  ;
      CLR   ;
      A     BR;
      )     ;
      JNB   M01b;
      L     DB7.DBW  444;
      T     DB3.DBB   64;
      SET   ;
      SAVE  ;
      CLR   ;
M01b: A     BR;
      )     ;
      JNB   M01c;
      L     DB7.DBW  446;
      T     DB3.DBB  101;
M01c: NOP   0;
NETWORK
TITLE =
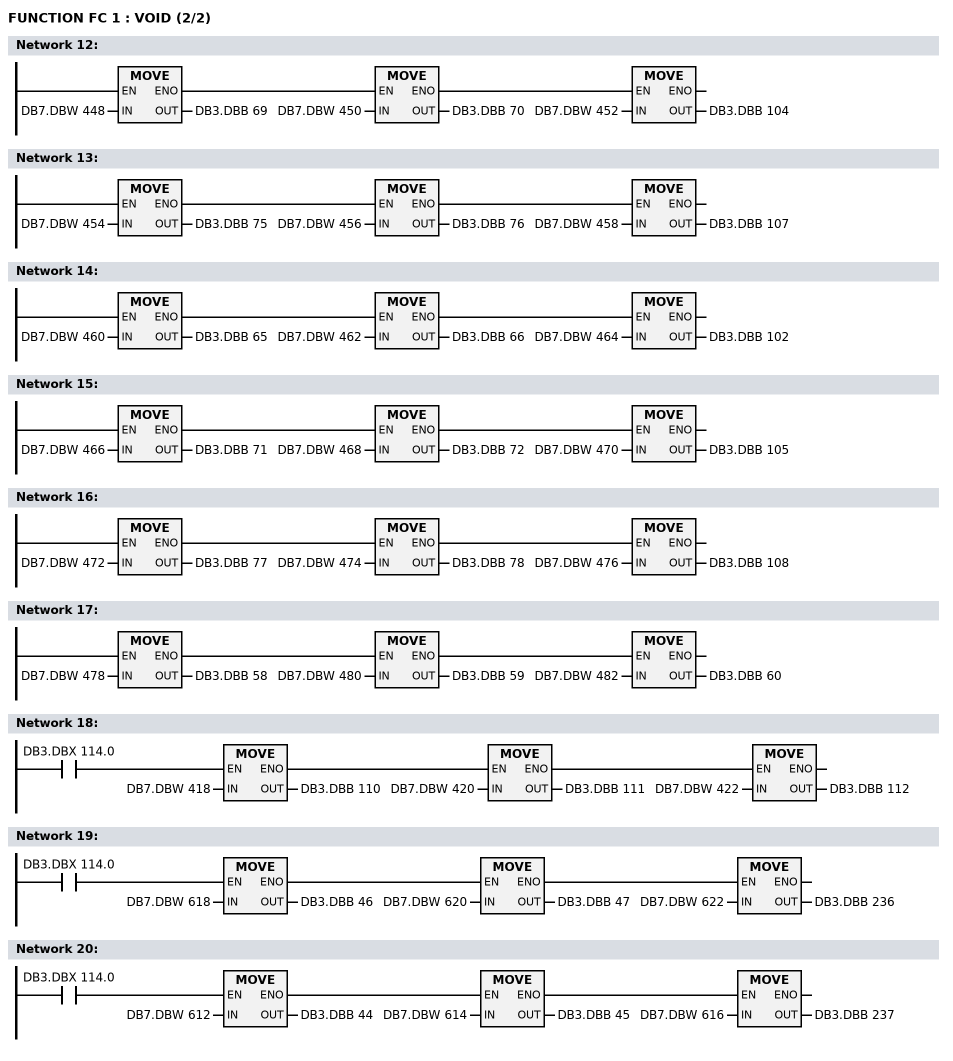

      A(    ;
      A(    ;
      L     DB7.DBW  448;
      T     DB3.DBB   69;
      SET   ;
      SAVE  ;
      CLR   ;
      A     BR;
      )     ;
      JNB   M01d;
      L     DB7.DBW  450;
      T     DB3.DBB   70;
      SET   ;
      SAVE  ;
      CLR   ;
M01d: A     BR;
      )     ;
      JNB   M01e;
      L     DB7.DBW  452;
      T     DB3.DBB  104;
M01e: NOP   0;
NETWORK
TITLE =

      A(    ;
      A(    ;
      L     DB7.DBW  454;
      T     DB3.DBB   75;
      SET   ;
      SAVE  ;
      CLR   ;
      A     BR;
      )     ;
      JNB   M01f;
      L     DB7.DBW  456;
      T     DB3.DBB   76;
      SET   ;
      SAVE  ;
      CLR   ;
M01f: A     BR;
      )     ;
      JNB   M020;
      L     DB7.DBW  458;
      T     DB3.DBB  107;
M020: NOP   0;
NETWORK
TITLE =

      A(    ;
      A(    ;
      L     DB7.DBW  460;
      T     DB3.DBB   65;
      SET   ;
      SAVE  ;
      CLR   ;
      A     BR;
      )     ;
      JNB   M021;
      L     DB7.DBW  462;
      T     DB3.DBB   66;
      SET   ;
      SAVE  ;
      CLR   ;
M021: A     BR;
      )     ;
      JNB   M022;
      L     DB7.DBW  464;
      T     DB3.DBB  102;
M022: NOP   0;
NETWORK
TITLE =

      A(    ;
      A(    ;
      L     DB7.DBW  466;
      T     DB3.DBB   71;
      SET   ;
      SAVE  ;
      CLR   ;
      A     BR;
      )     ;
      JNB   M023;
      L     DB7.DBW  468;
      T     DB3.DBB   72;
      SET   ;
      SAVE  ;
      CLR   ;
M023: A     BR;
      )     ;
      JNB   M024;
      L     DB7.DBW  470;
      T     DB3.DBB  105;
M024: NOP   0;
NETWORK
TITLE =

      A(    ;
      A(    ;
      L     DB7.DBW  472;
      T     DB3.DBB   77;
      SET   ;
      SAVE  ;
      CLR   ;
      A     BR;
      )     ;
      JNB   M025;
      L     DB7.DBW  474;
      T     DB3.DBB   78;
      SET   ;
      SAVE  ;
      CLR   ;
M025: A     BR;
      )     ;
      JNB   M00a;
      L     DB7.DBW  476;
      T     DB3.DBB  108;
M00a: NOP   0;
NETWORK
TITLE =

      A(    ;
      A(    ;
      L     DB7.DBW  478;
      T     DB3.DBB   58;
      SET   ;
      SAVE  ;
      CLR   ;
      A     BR;
      )     ;
      JNB   M00b;
      L     DB7.DBW  480;
      T     DB3.DBB   59;
      SET   ;
      SAVE  ;
      CLR   ;
M00b: A     BR;
      )     ;
      JNB   M00c;
      L     DB7.DBW  482;
      T     DB3.DBB   60;
M00c: NOP   0;
NETWORK
TITLE =

      A(    ;
      A(    ;
      A     DB3.DBX  114.0;
      JNB   M00d;
      L     DB7.DBW  418;
      T     DB3.DBB  110;
      SET   ;
      SAVE  ;
      CLR   ;
M00d: A     BR;
      )     ;
      JNB   M026;
      L     DB7.DBW  420;
      T     DB3.DBB  111;
      SET   ;
      SAVE  ;
      CLR   ;
M026: A     BR;
      )     ;
      JNB   M027;
      L     DB7.DBW  422;
      T     DB3.DBB  112;
M027: NOP   0;
NETWORK
TITLE =

      A(    ;
      A(    ;
      A     DB3.DBX  114.0;
      JNB   M028;
      L     DB7.DBW  618;
      T     DB3.DBB   46;
      SET   ;
      SAVE  ;
      CLR   ;
M028: A     BR;
      )     ;
      JNB   M029;
      L     DB7.DBW  620;
      T     DB3.DBB   47;
      SET   ;
      SAVE  ;
      CLR   ;
M029: A     BR;
      )     ;
      JNB   M02a;
      L     DB7.DBW  622;
      T     DB3.DBB  236;
M02a: NOP   0;
NETWORK
TITLE =

      A(    ;
      A(    ;
      A     DB3.DBX  114.0;
      JNB   M02b;
      L     DB7.DBW  612;
      T     DB3.DBB   44;
      SET   ;
      SAVE  ;
      CLR   ;
M02b: A     BR;
      )     ;
      JNB   M02c;
      L     DB7.DBW  614;
      T     DB3.DBB   45;
      SET   ;
      SAVE  ;
      CLR   ;
M02c: A     BR;
      )     ;
      JNB   M02d;
      L     DB7.DBW  616;
      T     DB3.DBB  237;
M02d: NOP   0;
END_FUNCTION

FUNCTION FC 9 : VOID
VERSION : 0.1

BEGIN
NETWORK
TITLE =
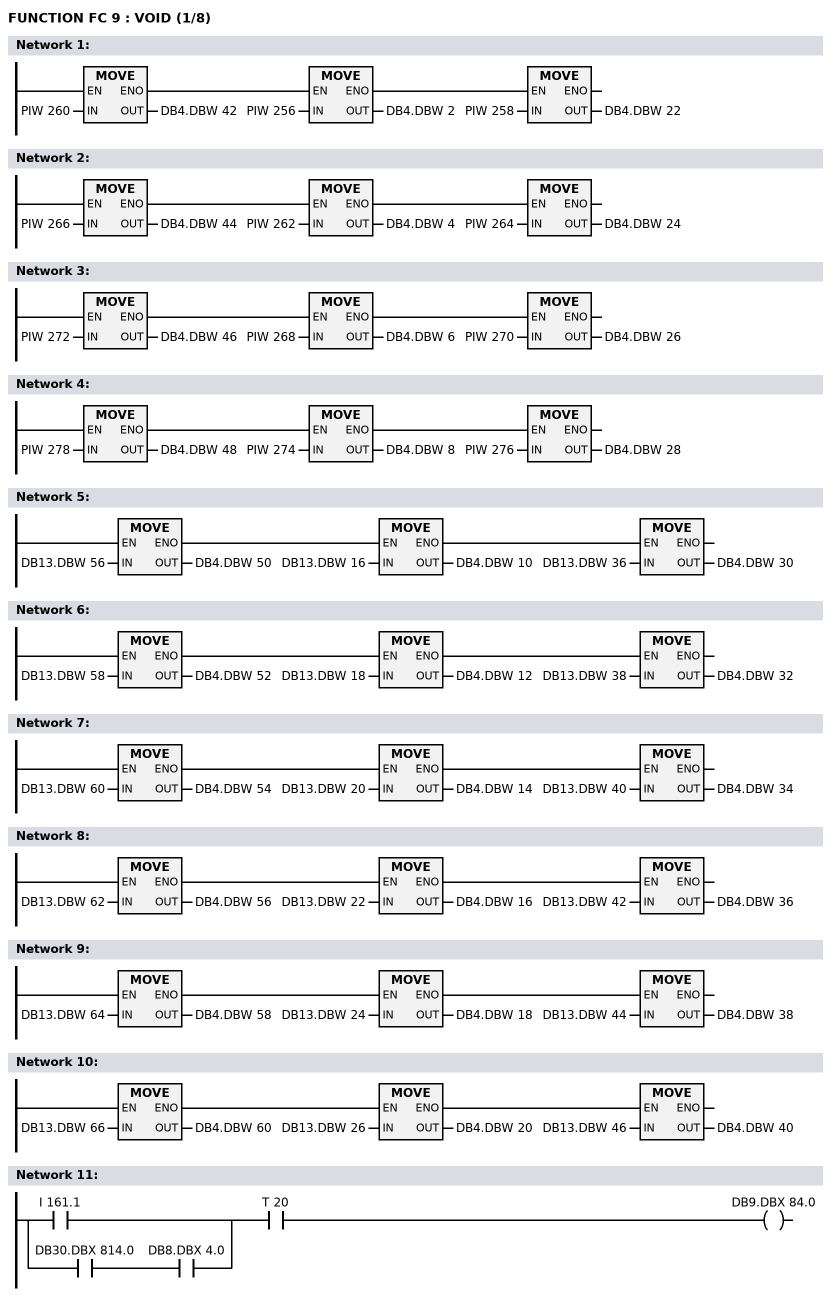

      A(    ;
      A(    ;
      L     PIW  260;
      T     DB4.DBW   42;
      SET   ;
      SAVE  ;
      CLR   ;
      A     BR;
      )     ;
      JNB   M001;
      L     PIW  256;
      T     DB4.DBW    2;
      SET   ;
      SAVE  ;
      CLR   ;
M001: A     BR;
      )     ;
      JNB   M002;
      L     PIW  258;
      T     DB4.DBW   22;
M002: NOP   0;
NETWORK
TITLE =

      A(    ;
      A(    ;
      L     PIW  266;
      T     DB4.DBW   44;
      SET   ;
      SAVE  ;
      CLR   ;
      A     BR;
      )     ;
      JNB   M003;
      L     PIW  262;
      T     DB4.DBW    4;
      SET   ;
      SAVE  ;
      CLR   ;
M003: A     BR;
      )     ;
      JNB   M004;
      L     PIW  264;
      T     DB4.DBW   24;
M004: NOP   0;
NETWORK
TITLE =

      A(    ;
      A(    ;
      L     PIW  272;
      T     DB4.DBW   46;
      SET   ;
      SAVE  ;
      CLR   ;
      A     BR;
      )     ;
      JNB   M005;
      L     PIW  268;
      T     DB4.DBW    6;
      SET   ;
      SAVE  ;
      CLR   ;
M005: A     BR;
      )     ;
      JNB   M006;
      L     PIW  270;
      T     DB4.DBW   26;
M006: NOP   0;
NETWORK
TITLE =

      A(    ;
      A(    ;
      L     PIW  278;
      T     DB4.DBW   48;
      SET   ;
      SAVE  ;
      CLR   ;
      A     BR;
      )     ;
      JNB   M007;
      L     PIW  274;
      T     DB4.DBW    8;
      SET   ;
      SAVE  ;
      CLR   ;
M007: A     BR;
      )     ;
      JNB   M008;
      L     PIW  276;
      T     DB4.DBW   28;
M008: NOP   0;
NETWORK
TITLE =

      A(    ;
      A(    ;
      L     DB13.DBW   56;
      T     DB4.DBW   50;
      SET   ;
      SAVE  ;
      CLR   ;
      A     BR;
      )     ;
      JNB   M009;
      L     DB13.DBW   16;
      T     DB4.DBW   10;
      SET   ;
      SAVE  ;
      CLR   ;
M009: A     BR;
      )     ;
      JNB   M00a;
      L     DB13.DBW   36;
      T     DB4.DBW   30;
M00a: NOP   0;
NETWORK
TITLE =

      A(    ;
      A(    ;
      L     DB13.DBW   58;
      T     DB4.DBW   52;
      SET   ;
      SAVE  ;
      CLR   ;
      A     BR;
      )     ;
      JNB   M00b;
      L     DB13.DBW   18;
      T     DB4.DBW   12;
      SET   ;
      SAVE  ;
      CLR   ;
M00b: A     BR;
      )     ;
      JNB   M00c;
      L     DB13.DBW   38;
      T     DB4.DBW   32;
M00c: NOP   0;
NETWORK
TITLE =

      A(    ;
      A(    ;
      L     DB13.DBW   60;
      T     DB4.DBW   54;
      SET   ;
      SAVE  ;
      CLR   ;
      A     BR;
      )     ;
      JNB   M00d;
      L     DB13.DBW   20;
      T     DB4.DBW   14;
      SET   ;
      SAVE  ;
      CLR   ;
M00d: A     BR;
      )     ;
      JNB   M00e;
      L     DB13.DBW   40;
      T     DB4.DBW   34;
M00e: NOP   0;
NETWORK
TITLE =

      A(    ;
      A(    ;
      L     DB13.DBW   62;
      T     DB4.DBW   56;
      SET   ;
      SAVE  ;
      CLR   ;
      A     BR;
      )     ;
      JNB   M00f;
      L     DB13.DBW   22;
      T     DB4.DBW   16;
      SET   ;
      SAVE  ;
      CLR   ;
M00f: A     BR;
      )     ;
      JNB   M010;
      L     DB13.DBW   42;
      T     DB4.DBW   36;
M010: NOP   0;
NETWORK
TITLE =

      A(    ;
      A(    ;
      L     DB13.DBW   64;
      T     DB4.DBW   58;
      SET   ;
      SAVE  ;
      CLR   ;
      A     BR;
      )     ;
      JNB   M011;
      L     DB13.DBW   24;
      T     DB4.DBW   18;
      SET   ;
      SAVE  ;
      CLR   ;
M011: A     BR;
      )     ;
      JNB   M012;
      L     DB13.DBW   44;
      T     DB4.DBW   38;
M012: NOP   0;
NETWORK
TITLE =

      A(    ;
      A(    ;
      L     DB13.DBW   66;
      T     DB4.DBW   60;
      SET   ;
      SAVE  ;
      CLR   ;
      A     BR;
      )     ;
      JNB   M013;
      L     DB13.DBW   26;
      T     DB4.DBW   20;
      SET   ;
      SAVE  ;
      CLR   ;
M013: A     BR;
      )     ;
      JNB   M014;
      L     DB13.DBW   46;
      T     DB4.DBW   40;
M014: NOP   0;
NETWORK
TITLE =

      A(    ;
      O     I    161.1;
      O     ;
      A     DB30.DBX  814.0;
      A     DB8.DBX    4.0;
      )     ;
      A     T     20;
      =     DB9.DBX   84.0;
NETWORK
TITLE =
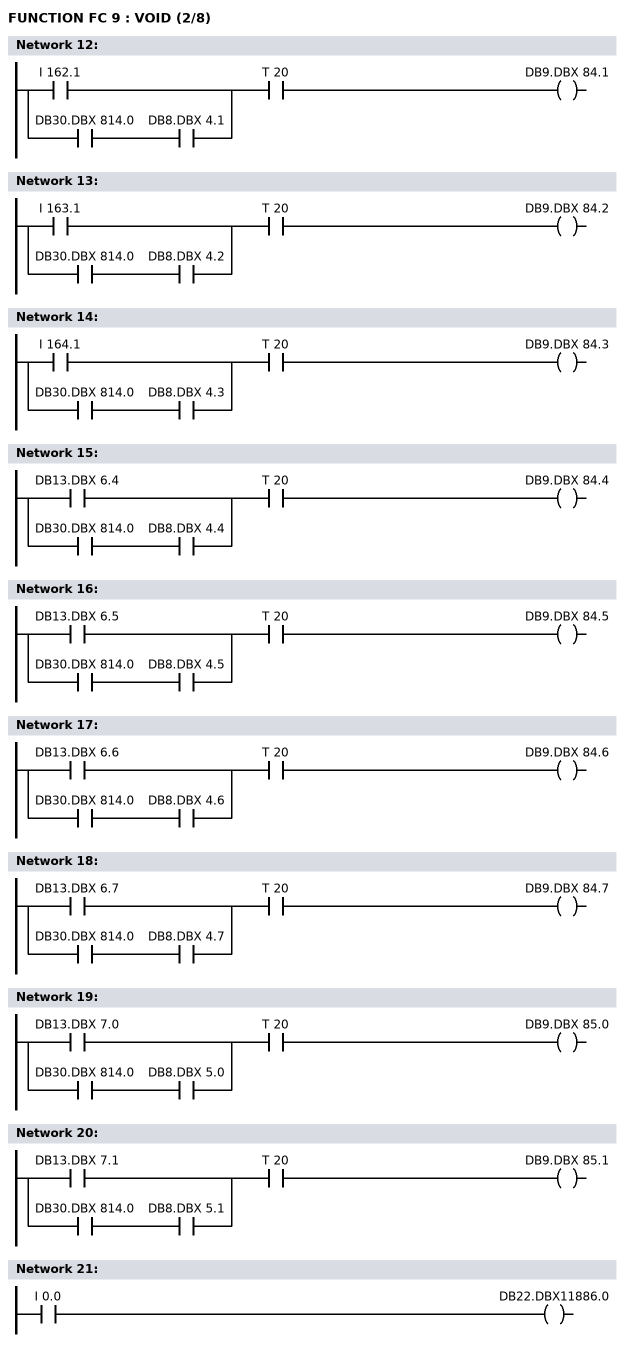

      A(    ;
      O     I    162.1;
      O     ;
      A     DB30.DBX  814.0;
      A     DB8.DBX    4.1;
      )     ;
      A     T     20;
      =     DB9.DBX   84.1;
NETWORK
TITLE =

      A(    ;
      O     I    163.1;
      O     ;
      A     DB30.DBX  814.0;
      A     DB8.DBX    4.2;
      )     ;
      A     T     20;
      =     DB9.DBX   84.2;
NETWORK
TITLE =

      A(    ;
      O     I    164.1;
      O     ;
      A     DB30.DBX  814.0;
      A     DB8.DBX    4.3;
      )     ;
      A     T     20;
      =     DB9.DBX   84.3;
NETWORK
TITLE =

      A(    ;
      O     DB13.DBX    6.4;
      O     ;
      A     DB30.DBX  814.0;
      A     DB8.DBX    4.4;
      )     ;
      A     T     20;
      =     DB9.DBX   84.4;
NETWORK
TITLE =

      A(    ;
      O     DB13.DBX    6.5;
      O     ;
      A     DB30.DBX  814.0;
      A     DB8.DBX    4.5;
      )     ;
      A     T     20;
      =     DB9.DBX   84.5;
NETWORK
TITLE =

      A(    ;
      O     DB13.DBX    6.6;
      O     ;
      A     DB30.DBX  814.0;
      A     DB8.DBX    4.6;
      )     ;
      A     T     20;
      =     DB9.DBX   84.6;
NETWORK
TITLE =

      A(    ;
      O     DB13.DBX    6.7;
      O     ;
      A     DB30.DBX  814.0;
      A     DB8.DBX    4.7;
      )     ;
      A     T     20;
      =     DB9.DBX   84.7;
NETWORK
TITLE =

      A(    ;
      O     DB13.DBX    7.0;
      O     ;
      A     DB30.DBX  814.0;
      A     DB8.DBX    5.0;
      )     ;
      A     T     20;
      =     DB9.DBX   85.0;
NETWORK
TITLE =

      A(    ;
      O     DB13.DBX    7.1;
      O     ;
      A     DB30.DBX  814.0;
      A     DB8.DBX    5.1;
      )     ;
      A     T     20;
      =     DB9.DBX   85.1;
NETWORK
TITLE =

      A     I      0.0;
      =     DB22.DBX11886.0;
NETWORK
TITLE =
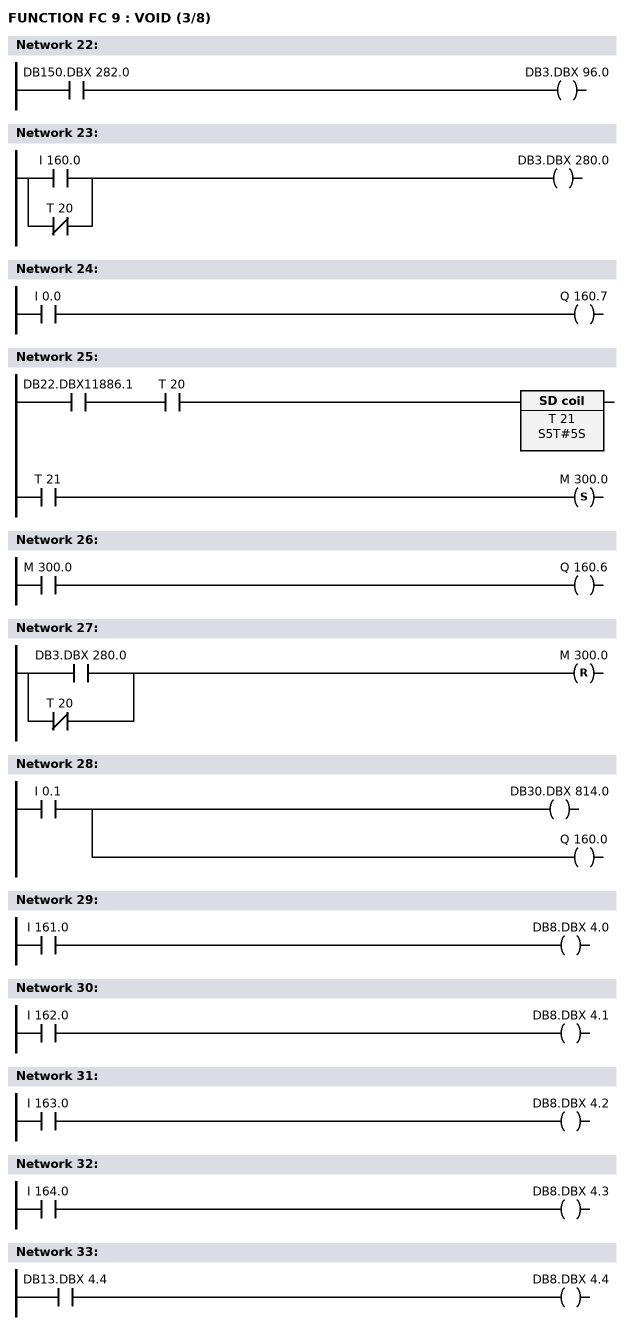

      A     DB150.DBX  282.0;
      =     DB3.DBX   96.0;
NETWORK
TITLE =

      O     I    160.0;
      ON    T     20;
      =     DB3.DBX  280.0;
NETWORK
TITLE =

      A     I      0.0;
      =     Q    160.7;
NETWORK
TITLE =

      A     DB22.DBX11886.1;
      A     T     20;
      L     S5T#5S;
      SD    T     21;
      NOP   0;
      NOP   0;
      NOP   0;
      A     T     21;
      S     M    300.0;
NETWORK
TITLE =

      A     M    300.0;
      =     Q    160.6;
NETWORK
TITLE =

      O     DB3.DBX  280.0;
      ON    T     20;
      R     M    300.0;
NETWORK
TITLE =

      A     I      0.1;
      =     DB30.DBX  814.0;
      =     Q    160.0;
NETWORK
TITLE =

      A     I    161.0;
      =     DB8.DBX    4.0;
NETWORK
TITLE =

      A     I    162.0;
      =     DB8.DBX    4.1;
NETWORK
TITLE =

      A     I    163.0;
      =     DB8.DBX    4.2;
NETWORK
TITLE =

      A     I    164.0;
      =     DB8.DBX    4.3;
NETWORK
TITLE =

      A     DB13.DBX    4.4;
      =     DB8.DBX    4.4;
NETWORK
TITLE =
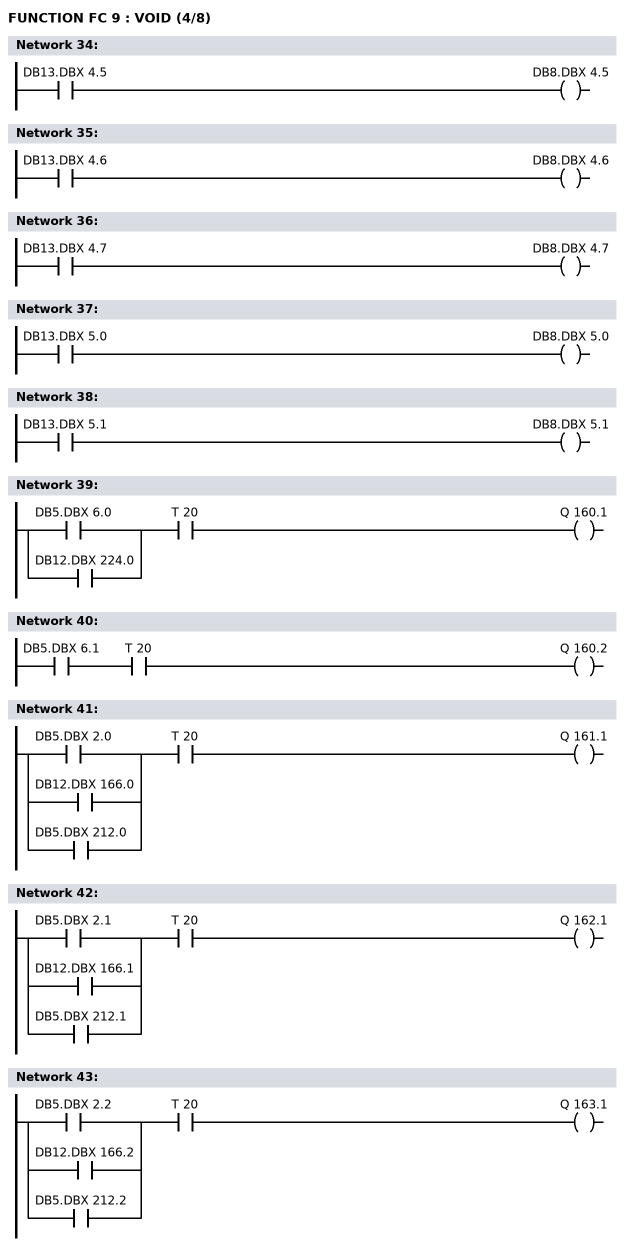

      A     DB13.DBX    4.5;
      =     DB8.DBX    4.5;
NETWORK
TITLE =

      A     DB13.DBX    4.6;
      =     DB8.DBX    4.6;
NETWORK
TITLE =

      A     DB13.DBX    4.7;
      =     DB8.DBX    4.7;
NETWORK
TITLE =

      A     DB13.DBX    5.0;
      =     DB8.DBX    5.0;
NETWORK
TITLE =

      A     DB13.DBX    5.1;
      =     DB8.DBX    5.1;
NETWORK
TITLE =

      A(    ;
      O     DB5.DBX    6.0;
      O     DB12.DBX  224.0;
      )     ;
      A     T     20;
      =     Q    160.1;
NETWORK
TITLE =

      A     DB5.DBX    6.1;
      A     T     20;
      =     Q    160.2;
NETWORK
TITLE =

      A(    ;
      O     DB5.DBX    2.0;
      O     DB12.DBX  166.0;
      O     DB5.DBX  212.0;
      )     ;
      A     T     20;
      =     Q    161.1;
NETWORK
TITLE =

      A(    ;
      O     DB5.DBX    2.1;
      O     DB12.DBX  166.1;
      O     DB5.DBX  212.1;
      )     ;
      A     T     20;
      =     Q    162.1;
NETWORK
TITLE =

      A(    ;
      O     DB5.DBX    2.2;
      O     DB12.DBX  166.2;
      O     DB5.DBX  212.2;
      )     ;
      A     T     20;
      =     Q    163.1;
NETWORK
TITLE =
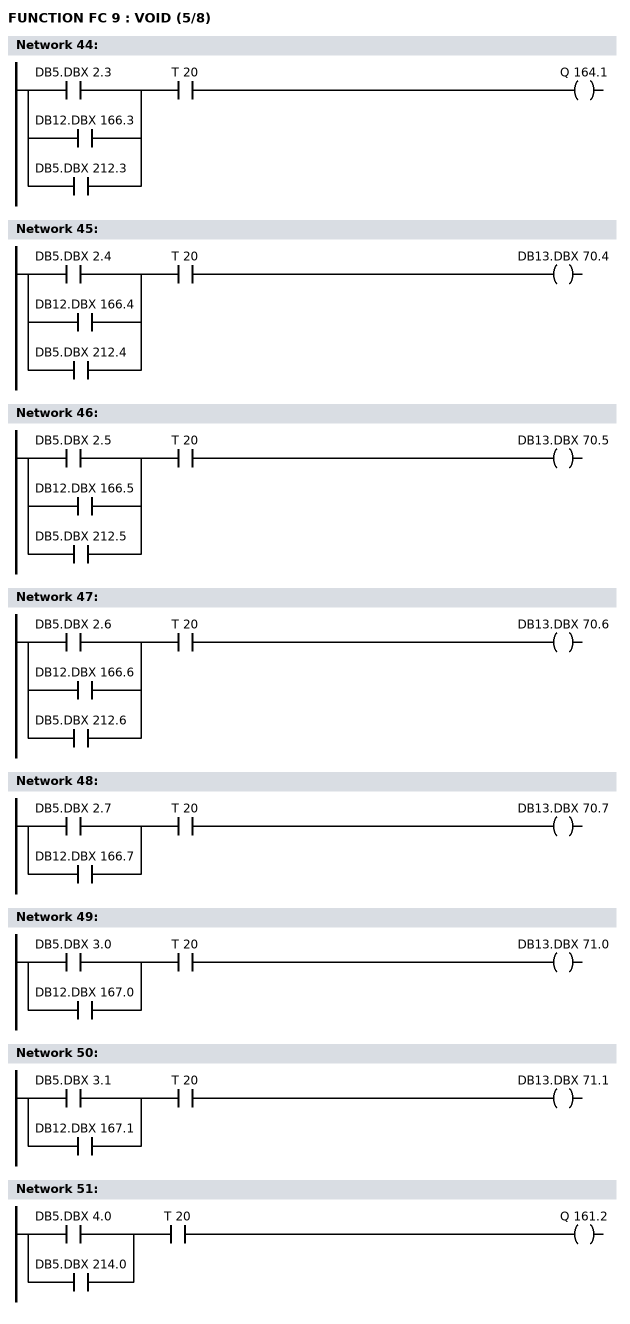

      A(    ;
      O     DB5.DBX    2.3;
      O     DB12.DBX  166.3;
      O     DB5.DBX  212.3;
      )     ;
      A     T     20;
      =     Q    164.1;
NETWORK
TITLE =

      A(    ;
      O     DB5.DBX    2.4;
      O     DB12.DBX  166.4;
      O     DB5.DBX  212.4;
      )     ;
      A     T     20;
      =     DB13.DBX   70.4;
NETWORK
TITLE =

      A(    ;
      O     DB5.DBX    2.5;
      O     DB12.DBX  166.5;
      O     DB5.DBX  212.5;
      )     ;
      A     T     20;
      =     DB13.DBX   70.5;
NETWORK
TITLE =

      A(    ;
      O     DB5.DBX    2.6;
      O     DB12.DBX  166.6;
      O     DB5.DBX  212.6;
      )     ;
      A     T     20;
      =     DB13.DBX   70.6;
NETWORK
TITLE =

      A(    ;
      O     DB5.DBX    2.7;
      O     DB12.DBX  166.7;
      )     ;
      A     T     20;
      =     DB13.DBX   70.7;
NETWORK
TITLE =

      A(    ;
      O     DB5.DBX    3.0;
      O     DB12.DBX  167.0;
      )     ;
      A     T     20;
      =     DB13.DBX   71.0;
NETWORK
TITLE =

      A(    ;
      O     DB5.DBX    3.1;
      O     DB12.DBX  167.1;
      )     ;
      A     T     20;
      =     DB13.DBX   71.1;
NETWORK
TITLE =

      A(    ;
      O     DB5.DBX    4.0;
      O     DB5.DBX  214.0;
      )     ;
      A     T     20;
      =     Q    161.2;
NETWORK
TITLE =
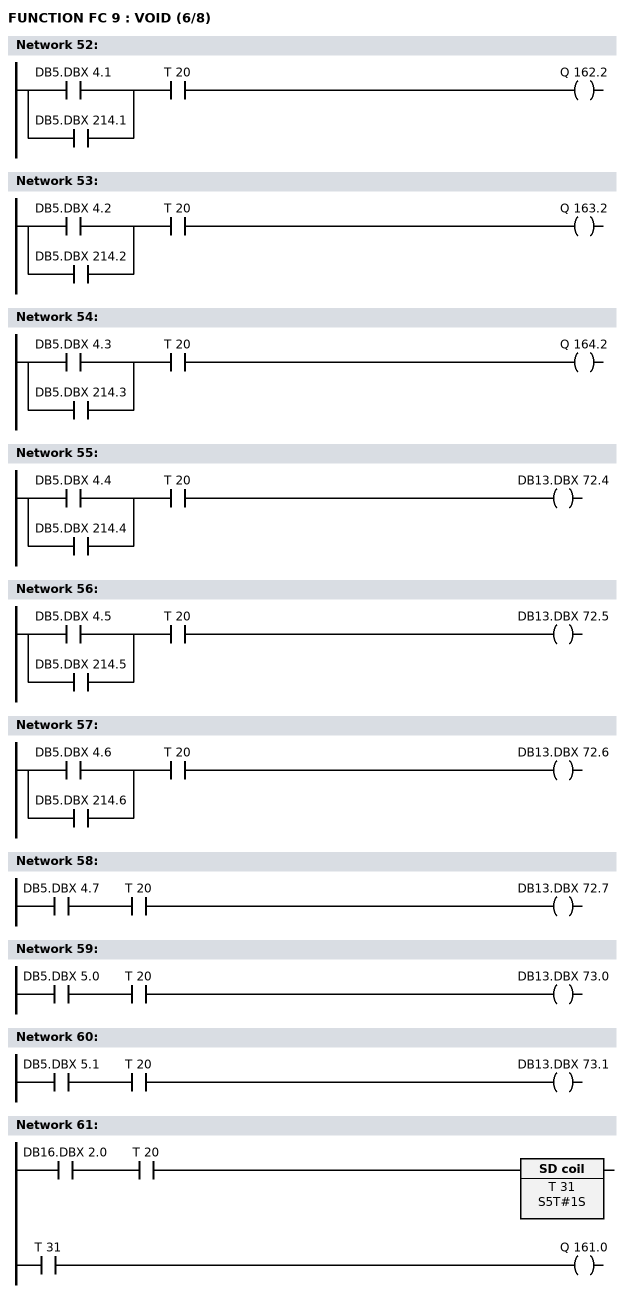

      A(    ;
      O     DB5.DBX    4.1;
      O     DB5.DBX  214.1;
      )     ;
      A     T     20;
      =     Q    162.2;
NETWORK
TITLE =

      A(    ;
      O     DB5.DBX    4.2;
      O     DB5.DBX  214.2;
      )     ;
      A     T     20;
      =     Q    163.2;
NETWORK
TITLE =

      A(    ;
      O     DB5.DBX    4.3;
      O     DB5.DBX  214.3;
      )     ;
      A     T     20;
      =     Q    164.2;
NETWORK
TITLE =

      A(    ;
      O     DB5.DBX    4.4;
      O     DB5.DBX  214.4;
      )     ;
      A     T     20;
      =     DB13.DBX   72.4;
NETWORK
TITLE =

      A(    ;
      O     DB5.DBX    4.5;
      O     DB5.DBX  214.5;
      )     ;
      A     T     20;
      =     DB13.DBX   72.5;
NETWORK
TITLE =

      A(    ;
      O     DB5.DBX    4.6;
      O     DB5.DBX  214.6;
      )     ;
      A     T     20;
      =     DB13.DBX   72.6;
NETWORK
TITLE =

      A     DB5.DBX    4.7;
      A     T     20;
      =     DB13.DBX   72.7;
NETWORK
TITLE =

      A     DB5.DBX    5.0;
      A     T     20;
      =     DB13.DBX   73.0;
NETWORK
TITLE =

      A     DB5.DBX    5.1;
      A     T     20;
      =     DB13.DBX   73.1;
NETWORK
TITLE =

      A     DB16.DBX    2.0;
      A     T     20;
      L     S5T#1S;
      SD    T     31;
      NOP   0;
      NOP   0;
      NOP   0;
      A     T     31;
      =     Q    161.0;
NETWORK
TITLE =
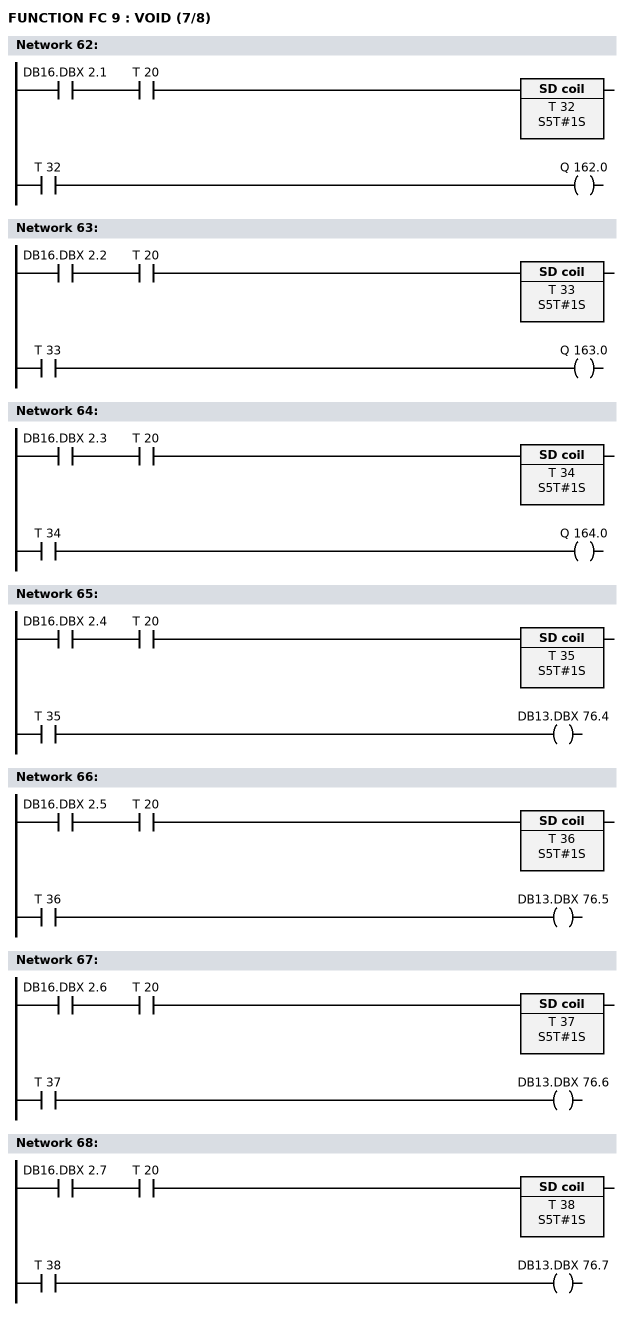

      A     DB16.DBX    2.1;
      A     T     20;
      L     S5T#1S;
      SD    T     32;
      NOP   0;
      NOP   0;
      NOP   0;
      A     T     32;
      =     Q    162.0;
NETWORK
TITLE =

      A     DB16.DBX    2.2;
      A     T     20;
      L     S5T#1S;
      SD    T     33;
      NOP   0;
      NOP   0;
      NOP   0;
      A     T     33;
      =     Q    163.0;
NETWORK
TITLE =

      A     DB16.DBX    2.3;
      A     T     20;
      L     S5T#1S;
      SD    T     34;
      NOP   0;
      NOP   0;
      NOP   0;
      A     T     34;
      =     Q    164.0;
NETWORK
TITLE =

      A     DB16.DBX    2.4;
      A     T     20;
      L     S5T#1S;
      SD    T     35;
      NOP   0;
      NOP   0;
      NOP   0;
      A     T     35;
      =     DB13.DBX   76.4;
NETWORK
TITLE =

      A     DB16.DBX    2.5;
      A     T     20;
      L     S5T#1S;
      SD    T     36;
      NOP   0;
      NOP   0;
      NOP   0;
      A     T     36;
      =     DB13.DBX   76.5;
NETWORK
TITLE =

      A     DB16.DBX    2.6;
      A     T     20;
      L     S5T#1S;
      SD    T     37;
      NOP   0;
      NOP   0;
      NOP   0;
      A     T     37;
      =     DB13.DBX   76.6;
NETWORK
TITLE =

      A     DB16.DBX    2.7;
      A     T     20;
      L     S5T#1S;
      SD    T     38;
      NOP   0;
      NOP   0;
      NOP   0;
      A     T     38;
      =     DB13.DBX   76.7;
NETWORK
TITLE =
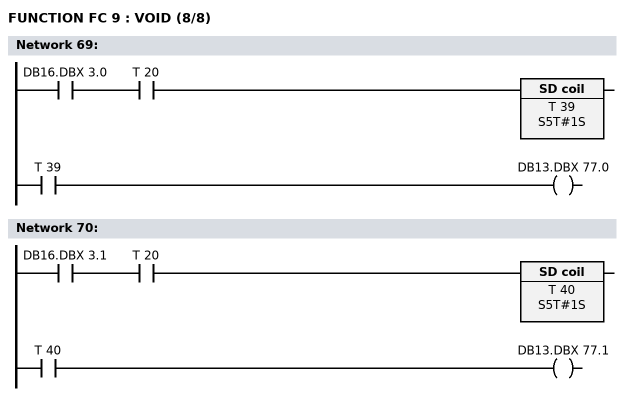

      A     DB16.DBX    3.0;
      A     T     20;
      L     S5T#1S;
      SD    T     39;
      NOP   0;
      NOP   0;
      NOP   0;
      A     T     39;
      =     DB13.DBX   77.0;
NETWORK
TITLE =

      A     DB16.DBX    3.1;
      A     T     20;
      L     S5T#1S;
      SD    T     40;
      NOP   0;
      NOP   0;
      NOP   0;
      A     T     40;
      =     DB13.DBX   77.1;
END_FUNCTION

FUNCTION FC 15 : VOID
VERSION : 0.1

BEGIN
NETWORK
TITLE =
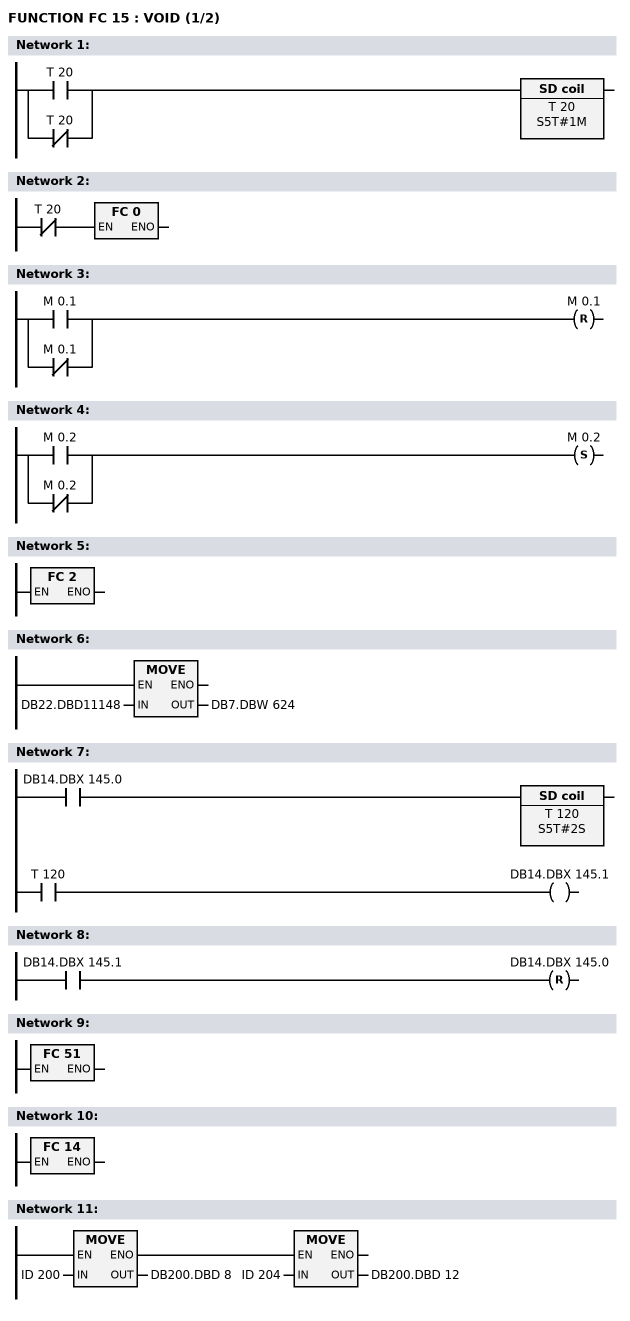

      A(    ;
      O     T     20;
      ON    T     20;
      )     ;
      L     S5T#1M;
      SD    T     20;
      NOP   0;
      NOP   0;
      NOP   0;
      NOP   0;
NETWORK
TITLE =

      AN    T     20;
      JNB   M002;
      CALL FC     0 ;
M002: NOP   0;
NETWORK
TITLE =

      O     M      0.1;
      ON    M      0.1;
      R     M      0.1;
NETWORK
TITLE =

      O     M      0.2;
      ON    M      0.2;
      S     M      0.2;
NETWORK
TITLE =

      CALL FC     2 ;
      NOP   0;
NETWORK
TITLE =

      L     DB22.DBD11148;
      T     DB7.DBW  624;
      NOP   0;
NETWORK
TITLE =

      A     DB14.DBX  145.0;
      L     S5T#2S;
      SD    T    120;
      NOP   0;
      NOP   0;
      NOP   0;
      A     T    120;
      =     DB14.DBX  145.1;
NETWORK
TITLE =

      A     DB14.DBX  145.1;
      R     DB14.DBX  145.0;
NETWORK
TITLE =

      CALL FC    51 ;
      NOP   0;
NETWORK
TITLE =

      CALL FC    14 ;
      NOP   0;
NETWORK
TITLE =

      A(    ;
      L     ID   200;
      T     DB200.DBD    8;
      SET   ;
      SAVE  ;
      CLR   ;
      A     BR;
      )     ;
      JNB   M003;
      L     ID   204;
      T     DB200.DBD   12;
M003: NOP   0;
NETWORK
TITLE =
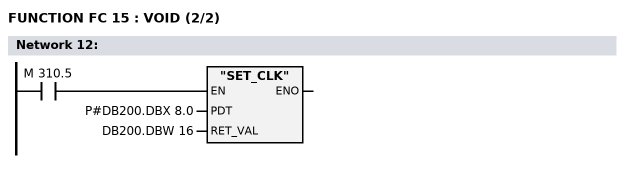

      A     M    310.5;
      JNB   M001;
      CALL "SET_CLK" (
           PDT                      := P#DB200.DBX 8.0,
           RET_VAL                  := DB200.DBW   16);
M001: NOP   0;
END_FUNCTION

FUNCTION FC 16 : VOID
VERSION : 0.1

BEGIN
NETWORK
TITLE =
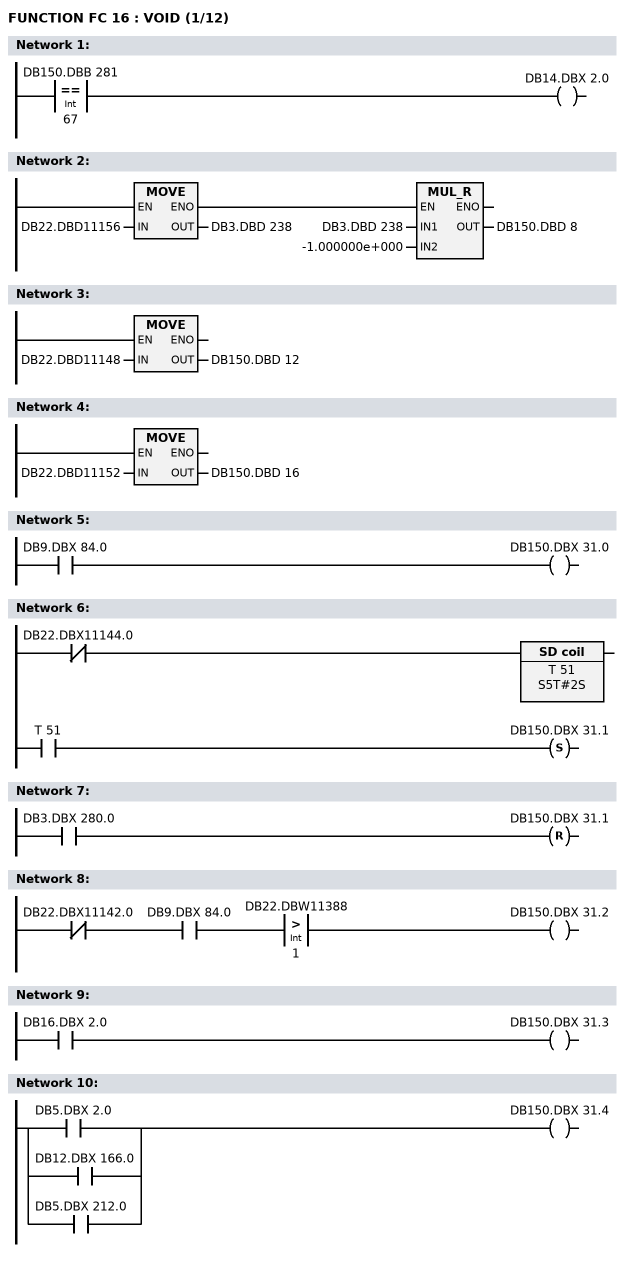

      L     DB150.DBB  281;
      L     67;
      ==I   ;
      =     DB14.DBX    2.0;
NETWORK
TITLE =

      A(    ;
      L     DB22.DBD11156;
      T     DB3.DBD  238;
      SET   ;
      SAVE  ;
      CLR   ;
      A     BR;
      )     ;
      JNB   M001;
      L     DB3.DBD  238;
      L     -1.000000e+000;
      *R    ;
      T     DB150.DBD    8;
M001: NOP   0;
NETWORK
TITLE =

      L     DB22.DBD11148;
      T     DB150.DBD   12;
      NOP   0;
NETWORK
TITLE =

      L     DB22.DBD11152;
      T     DB150.DBD   16;
      NOP   0;
NETWORK
TITLE =

      A     DB9.DBX   84.0;
      =     DB150.DBX   31.0;
NETWORK
TITLE =

      AN    DB22.DBX11144.0;
      L     S5T#2S;
      SD    T     51;
      NOP   0;
      NOP   0;
      NOP   0;
      A     T     51;
      S     DB150.DBX   31.1;
NETWORK
TITLE =

      A     DB3.DBX  280.0;
      R     DB150.DBX   31.1;
NETWORK
TITLE =

      AN    DB22.DBX11142.0;
      A     DB9.DBX   84.0;
      A(    ;
      L     DB22.DBW11388;
      L     1;
      >I    ;
      )     ;
      =     DB150.DBX   31.2;
NETWORK
TITLE =

      A     DB16.DBX    2.0;
      =     DB150.DBX   31.3;
NETWORK
TITLE =

      O     DB5.DBX    2.0;
      O     DB12.DBX  166.0;
      O     DB5.DBX  212.0;
      =     DB150.DBX   31.4;
NETWORK
TITLE =
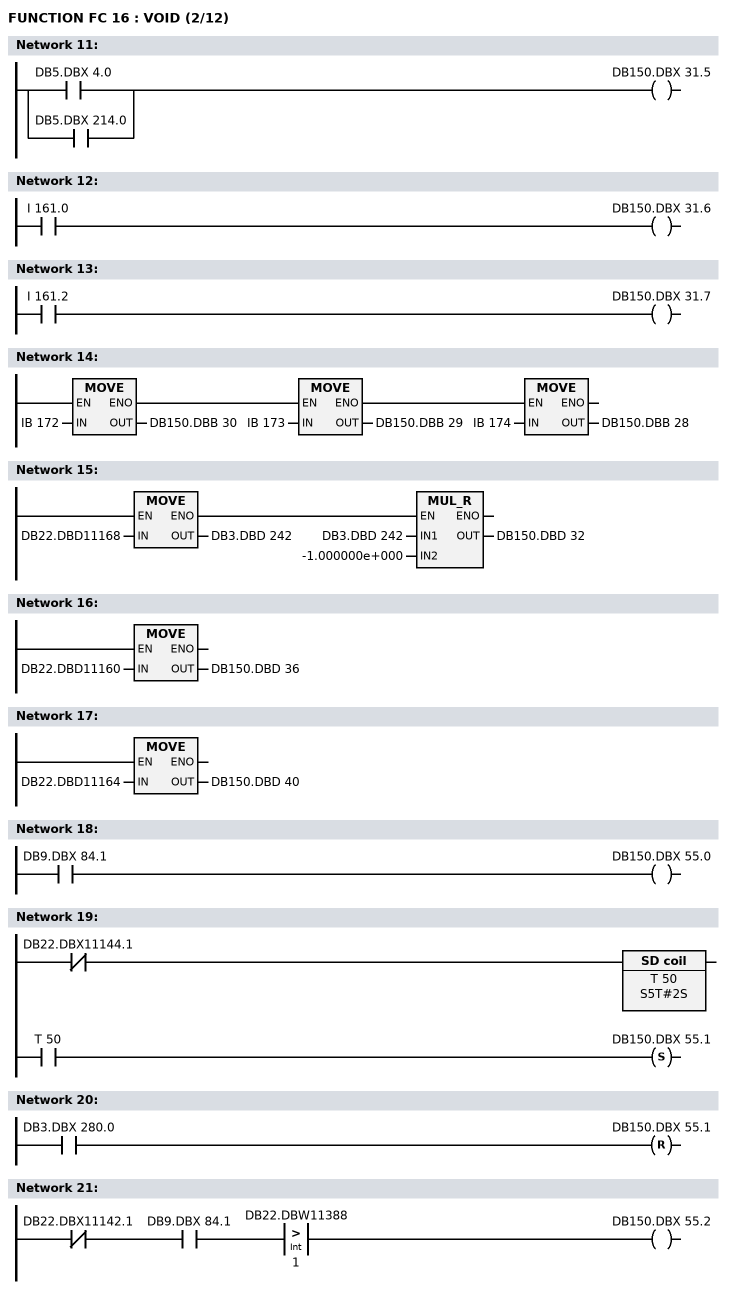

      O     DB5.DBX    4.0;
      O     DB5.DBX  214.0;
      =     DB150.DBX   31.5;
NETWORK
TITLE =

      A     I    161.0;
      =     DB150.DBX   31.6;
NETWORK
TITLE =

      A     I    161.2;
      =     DB150.DBX   31.7;
NETWORK
TITLE =

      A(    ;
      A(    ;
      L     IB   172;
      T     DB150.DBB   30;
      SET   ;
      SAVE  ;
      CLR   ;
      A     BR;
      )     ;
      JNB   M002;
      L     IB   173;
      T     DB150.DBB   29;
      SET   ;
      SAVE  ;
      CLR   ;
M002: A     BR;
      )     ;
      JNB   M003;
      L     IB   174;
      T     DB150.DBB   28;
M003: NOP   0;
NETWORK
TITLE =

      A(    ;
      L     DB22.DBD11168;
      T     DB3.DBD  242;
      SET   ;
      SAVE  ;
      CLR   ;
      A     BR;
      )     ;
      JNB   M004;
      L     DB3.DBD  242;
      L     -1.000000e+000;
      *R    ;
      T     DB150.DBD   32;
M004: NOP   0;
NETWORK
TITLE =

      L     DB22.DBD11160;
      T     DB150.DBD   36;
      NOP   0;
NETWORK
TITLE =

      L     DB22.DBD11164;
      T     DB150.DBD   40;
      NOP   0;
NETWORK
TITLE =

      A     DB9.DBX   84.1;
      =     DB150.DBX   55.0;
NETWORK
TITLE =

      AN    DB22.DBX11144.1;
      L     S5T#2S;
      SD    T     50;
      NOP   0;
      NOP   0;
      NOP   0;
      A     T     50;
      S     DB150.DBX   55.1;
NETWORK
TITLE =

      A     DB3.DBX  280.0;
      R     DB150.DBX   55.1;
NETWORK
TITLE =

      AN    DB22.DBX11142.1;
      A     DB9.DBX   84.1;
      A(    ;
      L     DB22.DBW11388;
      L     1;
      >I    ;
      )     ;
      =     DB150.DBX   55.2;
NETWORK
TITLE =
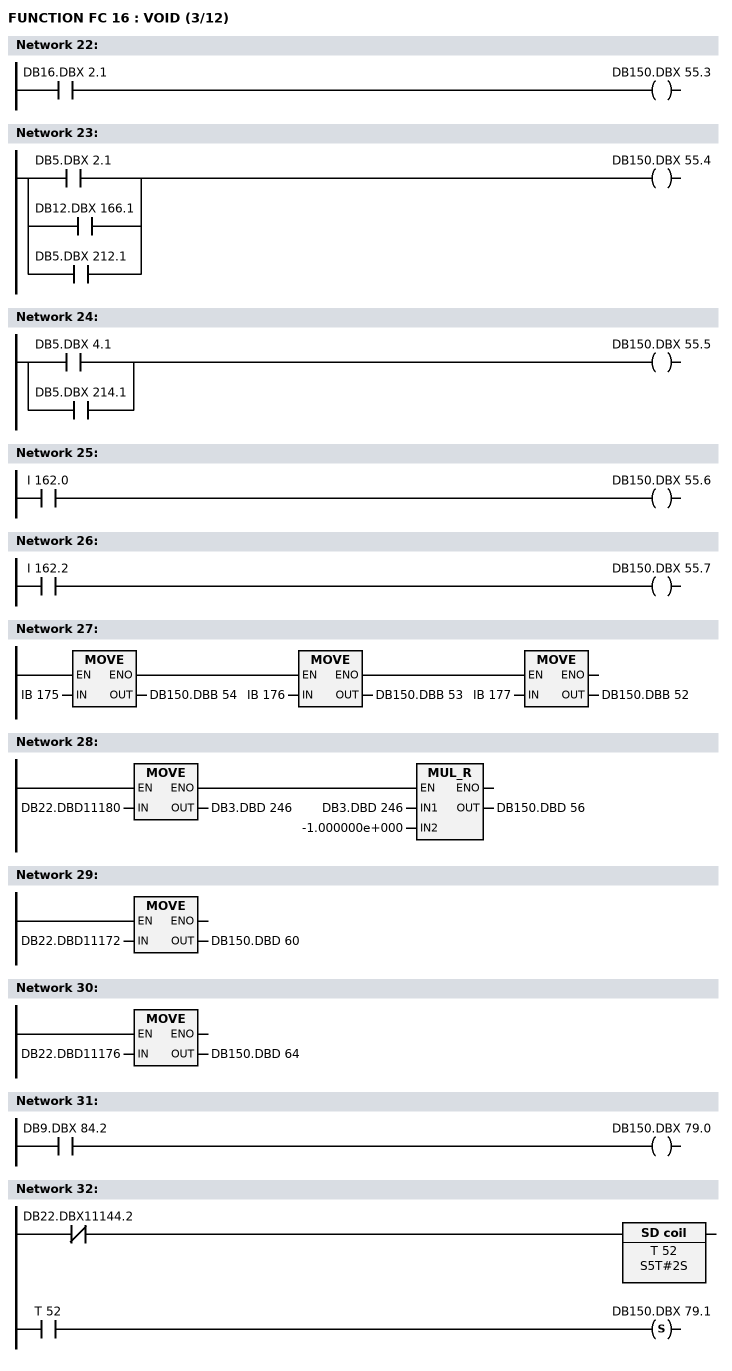

      A     DB16.DBX    2.1;
      =     DB150.DBX   55.3;
NETWORK
TITLE =

      O     DB5.DBX    2.1;
      O     DB12.DBX  166.1;
      O     DB5.DBX  212.1;
      =     DB150.DBX   55.4;
NETWORK
TITLE =

      O     DB5.DBX    4.1;
      O     DB5.DBX  214.1;
      =     DB150.DBX   55.5;
NETWORK
TITLE =

      A     I    162.0;
      =     DB150.DBX   55.6;
NETWORK
TITLE =

      A     I    162.2;
      =     DB150.DBX   55.7;
NETWORK
TITLE =

      A(    ;
      A(    ;
      L     IB   175;
      T     DB150.DBB   54;
      SET   ;
      SAVE  ;
      CLR   ;
      A     BR;
      )     ;
      JNB   M005;
      L     IB   176;
      T     DB150.DBB   53;
      SET   ;
      SAVE  ;
      CLR   ;
M005: A     BR;
      )     ;
      JNB   M006;
      L     IB   177;
      T     DB150.DBB   52;
M006: NOP   0;
NETWORK
TITLE =

      A(    ;
      L     DB22.DBD11180;
      T     DB3.DBD  246;
      SET   ;
      SAVE  ;
      CLR   ;
      A     BR;
      )     ;
      JNB   M007;
      L     DB3.DBD  246;
      L     -1.000000e+000;
      *R    ;
      T     DB150.DBD   56;
M007: NOP   0;
NETWORK
TITLE =

      L     DB22.DBD11172;
      T     DB150.DBD   60;
      NOP   0;
NETWORK
TITLE =

      L     DB22.DBD11176;
      T     DB150.DBD   64;
      NOP   0;
NETWORK
TITLE =

      A     DB9.DBX   84.2;
      =     DB150.DBX   79.0;
NETWORK
TITLE =

      AN    DB22.DBX11144.2;
      L     S5T#2S;
      SD    T     52;
      NOP   0;
      NOP   0;
      NOP   0;
      A     T     52;
      S     DB150.DBX   79.1;
NETWORK
TITLE =
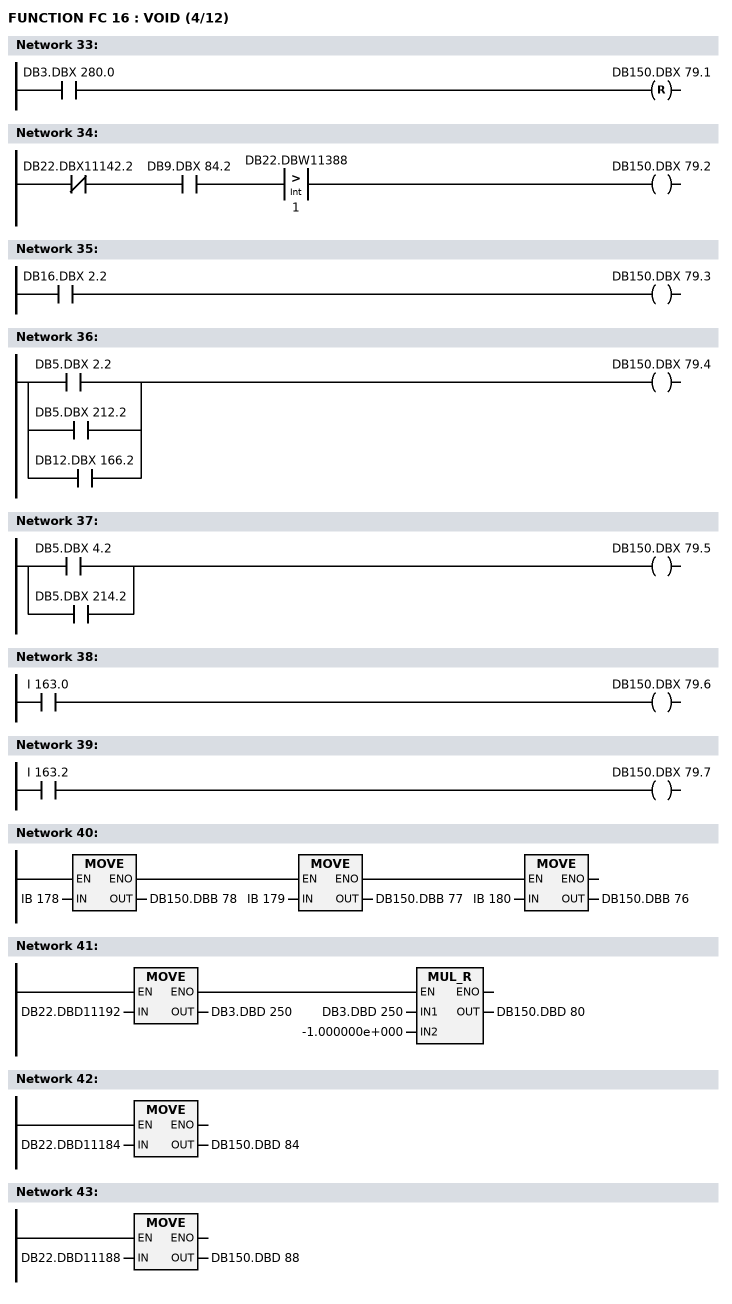

      A     DB3.DBX  280.0;
      R     DB150.DBX   79.1;
NETWORK
TITLE =

      AN    DB22.DBX11142.2;
      A     DB9.DBX   84.2;
      A(    ;
      L     DB22.DBW11388;
      L     1;
      >I    ;
      )     ;
      =     DB150.DBX   79.2;
NETWORK
TITLE =

      A     DB16.DBX    2.2;
      =     DB150.DBX   79.3;
NETWORK
TITLE =

      O     DB5.DBX    2.2;
      O     DB5.DBX  212.2;
      O     DB12.DBX  166.2;
      =     DB150.DBX   79.4;
NETWORK
TITLE =

      O     DB5.DBX    4.2;
      O     DB5.DBX  214.2;
      =     DB150.DBX   79.5;
NETWORK
TITLE =

      A     I    163.0;
      =     DB150.DBX   79.6;
NETWORK
TITLE =

      A     I    163.2;
      =     DB150.DBX   79.7;
NETWORK
TITLE =

      A(    ;
      A(    ;
      L     IB   178;
      T     DB150.DBB   78;
      SET   ;
      SAVE  ;
      CLR   ;
      A     BR;
      )     ;
      JNB   M008;
      L     IB   179;
      T     DB150.DBB   77;
      SET   ;
      SAVE  ;
      CLR   ;
M008: A     BR;
      )     ;
      JNB   M009;
      L     IB   180;
      T     DB150.DBB   76;
M009: NOP   0;
NETWORK
TITLE =

      A(    ;
      L     DB22.DBD11192;
      T     DB3.DBD  250;
      SET   ;
      SAVE  ;
      CLR   ;
      A     BR;
      )     ;
      JNB   M00a;
      L     DB3.DBD  250;
      L     -1.000000e+000;
      *R    ;
      T     DB150.DBD   80;
M00a: NOP   0;
NETWORK
TITLE =

      L     DB22.DBD11184;
      T     DB150.DBD   84;
      NOP   0;
NETWORK
TITLE =

      L     DB22.DBD11188;
      T     DB150.DBD   88;
      NOP   0;
NETWORK
TITLE =
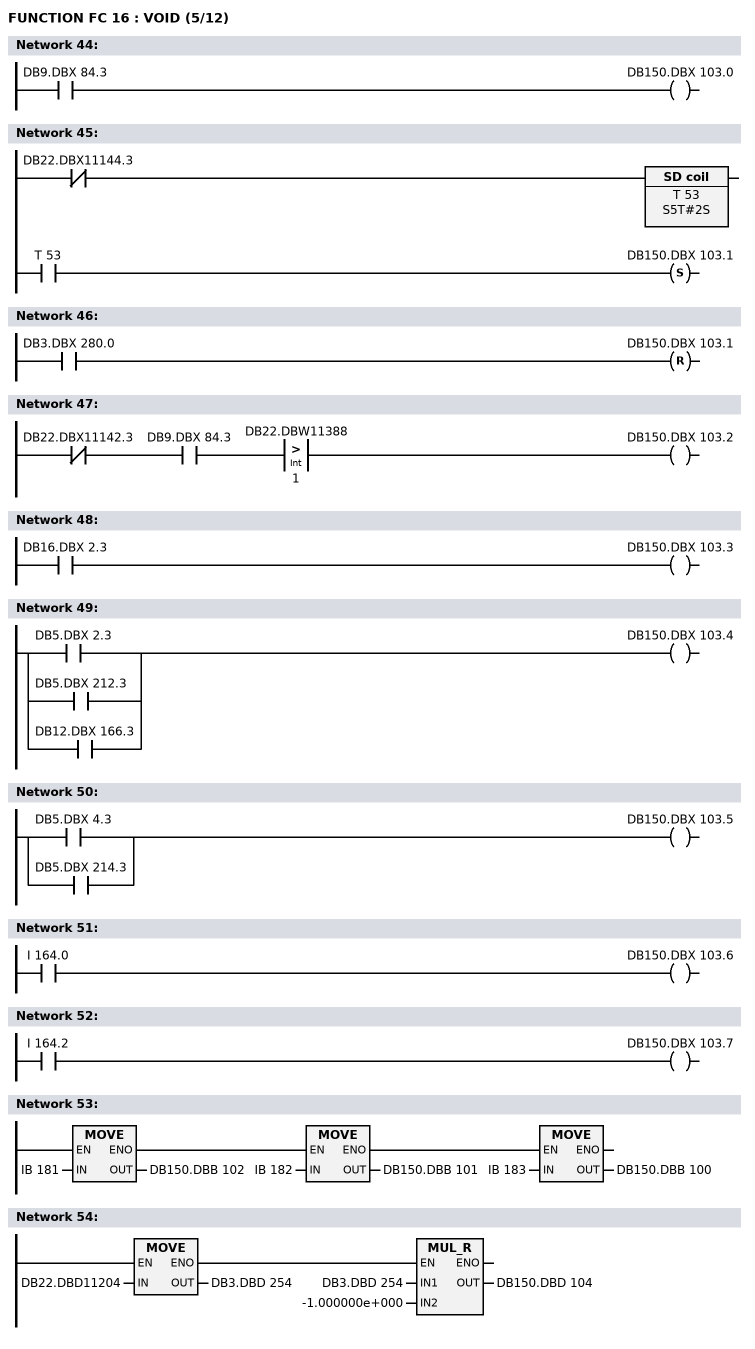

      A     DB9.DBX   84.3;
      =     DB150.DBX  103.0;
NETWORK
TITLE =

      AN    DB22.DBX11144.3;
      L     S5T#2S;
      SD    T     53;
      NOP   0;
      NOP   0;
      NOP   0;
      A     T     53;
      S     DB150.DBX  103.1;
NETWORK
TITLE =

      A     DB3.DBX  280.0;
      R     DB150.DBX  103.1;
NETWORK
TITLE =

      AN    DB22.DBX11142.3;
      A     DB9.DBX   84.3;
      A(    ;
      L     DB22.DBW11388;
      L     1;
      >I    ;
      )     ;
      =     DB150.DBX  103.2;
NETWORK
TITLE =

      A     DB16.DBX    2.3;
      =     DB150.DBX  103.3;
NETWORK
TITLE =

      O     DB5.DBX    2.3;
      O     DB5.DBX  212.3;
      O     DB12.DBX  166.3;
      =     DB150.DBX  103.4;
NETWORK
TITLE =

      O     DB5.DBX    4.3;
      O     DB5.DBX  214.3;
      =     DB150.DBX  103.5;
NETWORK
TITLE =

      A     I    164.0;
      =     DB150.DBX  103.6;
NETWORK
TITLE =

      A     I    164.2;
      =     DB150.DBX  103.7;
NETWORK
TITLE =

      A(    ;
      A(    ;
      L     IB   181;
      T     DB150.DBB  102;
      SET   ;
      SAVE  ;
      CLR   ;
      A     BR;
      )     ;
      JNB   M00b;
      L     IB   182;
      T     DB150.DBB  101;
      SET   ;
      SAVE  ;
      CLR   ;
M00b: A     BR;
      )     ;
      JNB   M00c;
      L     IB   183;
      T     DB150.DBB  100;
M00c: NOP   0;
NETWORK
TITLE =

      A(    ;
      L     DB22.DBD11204;
      T     DB3.DBD  254;
      SET   ;
      SAVE  ;
      CLR   ;
      A     BR;
      )     ;
      JNB   M00d;
      L     DB3.DBD  254;
      L     -1.000000e+000;
      *R    ;
      T     DB150.DBD  104;
M00d: NOP   0;
NETWORK
TITLE =
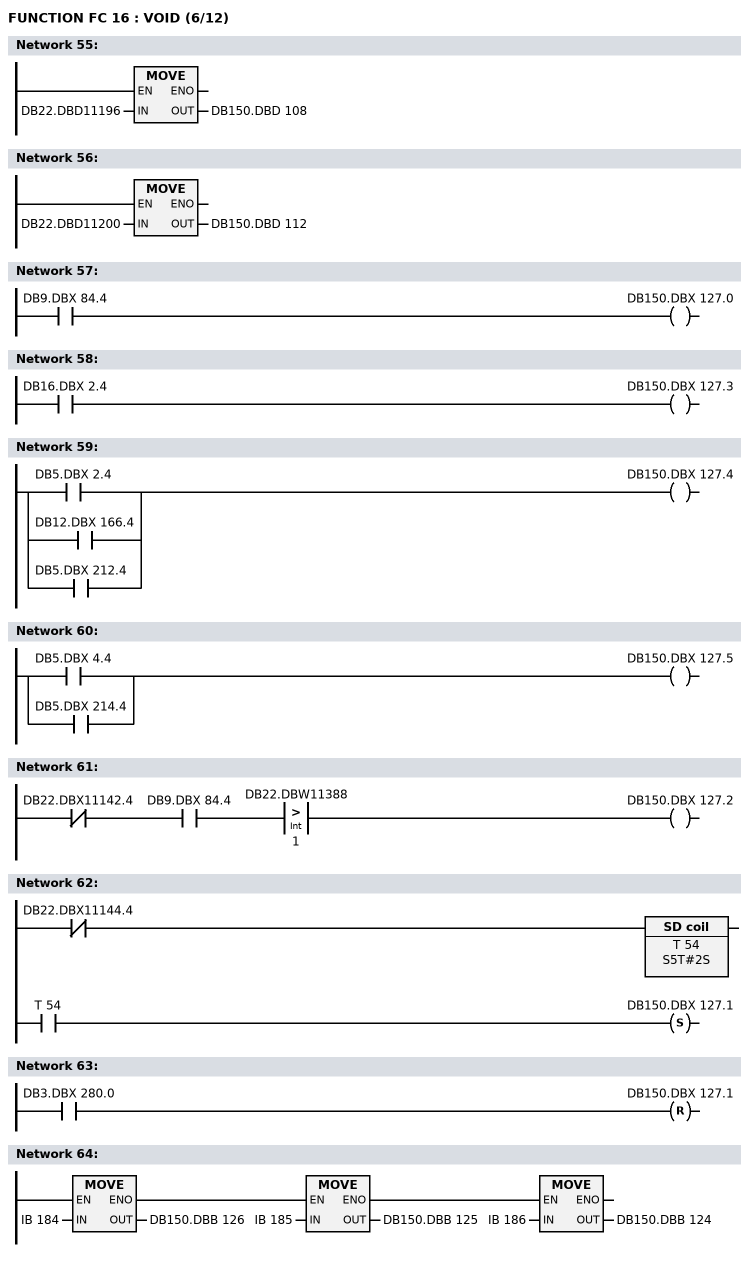

      L     DB22.DBD11196;
      T     DB150.DBD  108;
      NOP   0;
NETWORK
TITLE =

      L     DB22.DBD11200;
      T     DB150.DBD  112;
      NOP   0;
NETWORK
TITLE =

      A     DB9.DBX   84.4;
      =     DB150.DBX  127.0;
NETWORK
TITLE =

      A     DB16.DBX    2.4;
      =     DB150.DBX  127.3;
NETWORK
TITLE =

      O     DB5.DBX    2.4;
      O     DB12.DBX  166.4;
      O     DB5.DBX  212.4;
      =     DB150.DBX  127.4;
NETWORK
TITLE =

      O     DB5.DBX    4.4;
      O     DB5.DBX  214.4;
      =     DB150.DBX  127.5;
NETWORK
TITLE =

      AN    DB22.DBX11142.4;
      A     DB9.DBX   84.4;
      A(    ;
      L     DB22.DBW11388;
      L     1;
      >I    ;
      )     ;
      =     DB150.DBX  127.2;
NETWORK
TITLE =

      AN    DB22.DBX11144.4;
      L     S5T#2S;
      SD    T     54;
      NOP   0;
      NOP   0;
      NOP   0;
      A     T     54;
      S     DB150.DBX  127.1;
NETWORK
TITLE =

      A     DB3.DBX  280.0;
      R     DB150.DBX  127.1;
NETWORK
TITLE =

      A(    ;
      A(    ;
      L     IB   184;
      T     DB150.DBB  126;
      SET   ;
      SAVE  ;
      CLR   ;
      A     BR;
      )     ;
      JNB   M00e;
      L     IB   185;
      T     DB150.DBB  125;
      SET   ;
      SAVE  ;
      CLR   ;
M00e: A     BR;
      )     ;
      JNB   M00f;
      L     IB   186;
      T     DB150.DBB  124;
M00f: NOP   0;
NETWORK
TITLE =
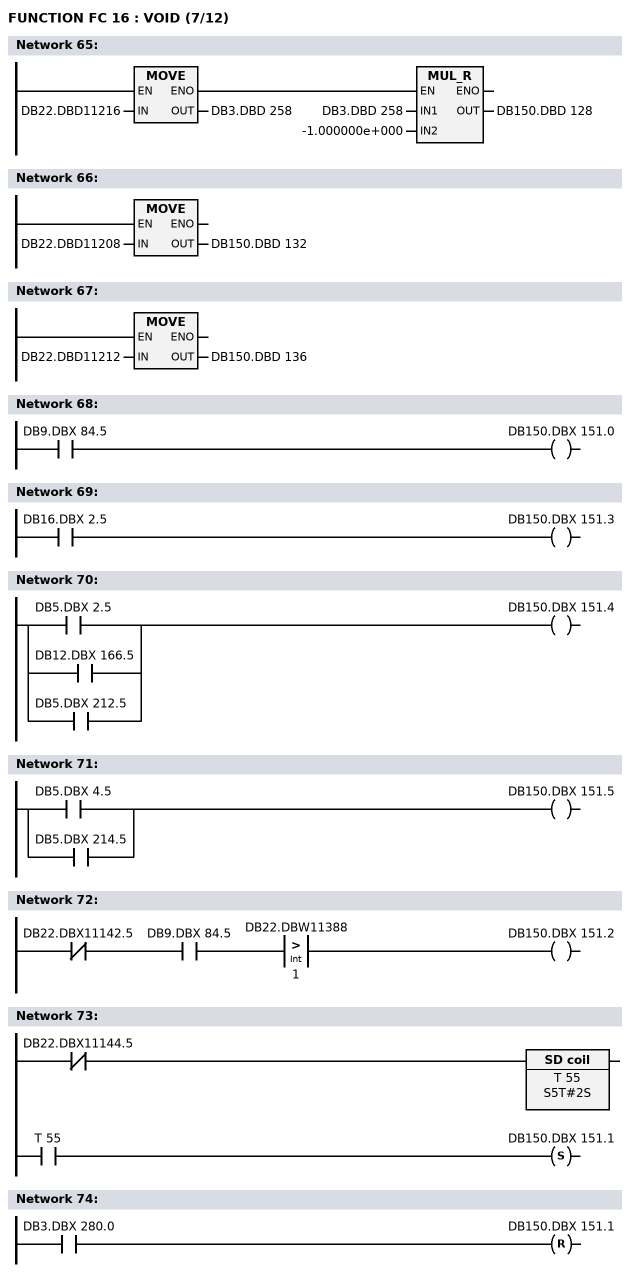

      A(    ;
      L     DB22.DBD11216;
      T     DB3.DBD  258;
      SET   ;
      SAVE  ;
      CLR   ;
      A     BR;
      )     ;
      JNB   M010;
      L     DB3.DBD  258;
      L     -1.000000e+000;
      *R    ;
      T     DB150.DBD  128;
M010: NOP   0;
NETWORK
TITLE =

      L     DB22.DBD11208;
      T     DB150.DBD  132;
      NOP   0;
NETWORK
TITLE =

      L     DB22.DBD11212;
      T     DB150.DBD  136;
      NOP   0;
NETWORK
TITLE =

      A     DB9.DBX   84.5;
      =     DB150.DBX  151.0;
NETWORK
TITLE =

      A     DB16.DBX    2.5;
      =     DB150.DBX  151.3;
NETWORK
TITLE =

      O     DB5.DBX    2.5;
      O     DB12.DBX  166.5;
      O     DB5.DBX  212.5;
      =     DB150.DBX  151.4;
NETWORK
TITLE =

      O     DB5.DBX    4.5;
      O     DB5.DBX  214.5;
      =     DB150.DBX  151.5;
NETWORK
TITLE =

      AN    DB22.DBX11142.5;
      A     DB9.DBX   84.5;
      A(    ;
      L     DB22.DBW11388;
      L     1;
      >I    ;
      )     ;
      =     DB150.DBX  151.2;
NETWORK
TITLE =

      AN    DB22.DBX11144.5;
      L     S5T#2S;
      SD    T     55;
      NOP   0;
      NOP   0;
      NOP   0;
      A     T     55;
      S     DB150.DBX  151.1;
NETWORK
TITLE =

      A     DB3.DBX  280.0;
      R     DB150.DBX  151.1;
NETWORK
TITLE =
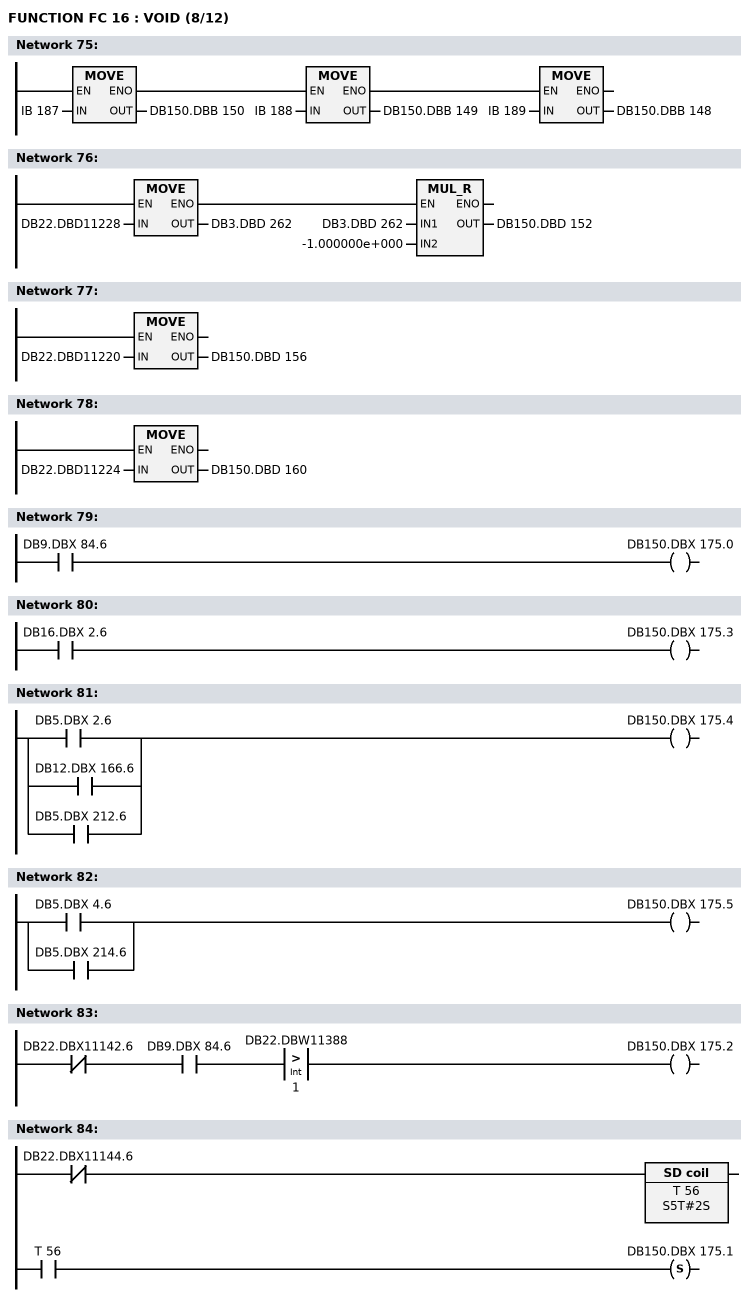

      A(    ;
      A(    ;
      L     IB   187;
      T     DB150.DBB  150;
      SET   ;
      SAVE  ;
      CLR   ;
      A     BR;
      )     ;
      JNB   M011;
      L     IB   188;
      T     DB150.DBB  149;
      SET   ;
      SAVE  ;
      CLR   ;
M011: A     BR;
      )     ;
      JNB   M012;
      L     IB   189;
      T     DB150.DBB  148;
M012: NOP   0;
NETWORK
TITLE =

      A(    ;
      L     DB22.DBD11228;
      T     DB3.DBD  262;
      SET   ;
      SAVE  ;
      CLR   ;
      A     BR;
      )     ;
      JNB   M013;
      L     DB3.DBD  262;
      L     -1.000000e+000;
      *R    ;
      T     DB150.DBD  152;
M013: NOP   0;
NETWORK
TITLE =

      L     DB22.DBD11220;
      T     DB150.DBD  156;
      NOP   0;
NETWORK
TITLE =

      L     DB22.DBD11224;
      T     DB150.DBD  160;
      NOP   0;
NETWORK
TITLE =

      A     DB9.DBX   84.6;
      =     DB150.DBX  175.0;
NETWORK
TITLE =

      A     DB16.DBX    2.6;
      =     DB150.DBX  175.3;
NETWORK
TITLE =

      O     DB5.DBX    2.6;
      O     DB12.DBX  166.6;
      O     DB5.DBX  212.6;
      =     DB150.DBX  175.4;
NETWORK
TITLE =

      O     DB5.DBX    4.6;
      O     DB5.DBX  214.6;
      =     DB150.DBX  175.5;
NETWORK
TITLE =

      AN    DB22.DBX11142.6;
      A     DB9.DBX   84.6;
      A(    ;
      L     DB22.DBW11388;
      L     1;
      >I    ;
      )     ;
      =     DB150.DBX  175.2;
NETWORK
TITLE =

      AN    DB22.DBX11144.6;
      L     S5T#2S;
      SD    T     56;
      NOP   0;
      NOP   0;
      NOP   0;
      A     T     56;
      S     DB150.DBX  175.1;
NETWORK
TITLE =
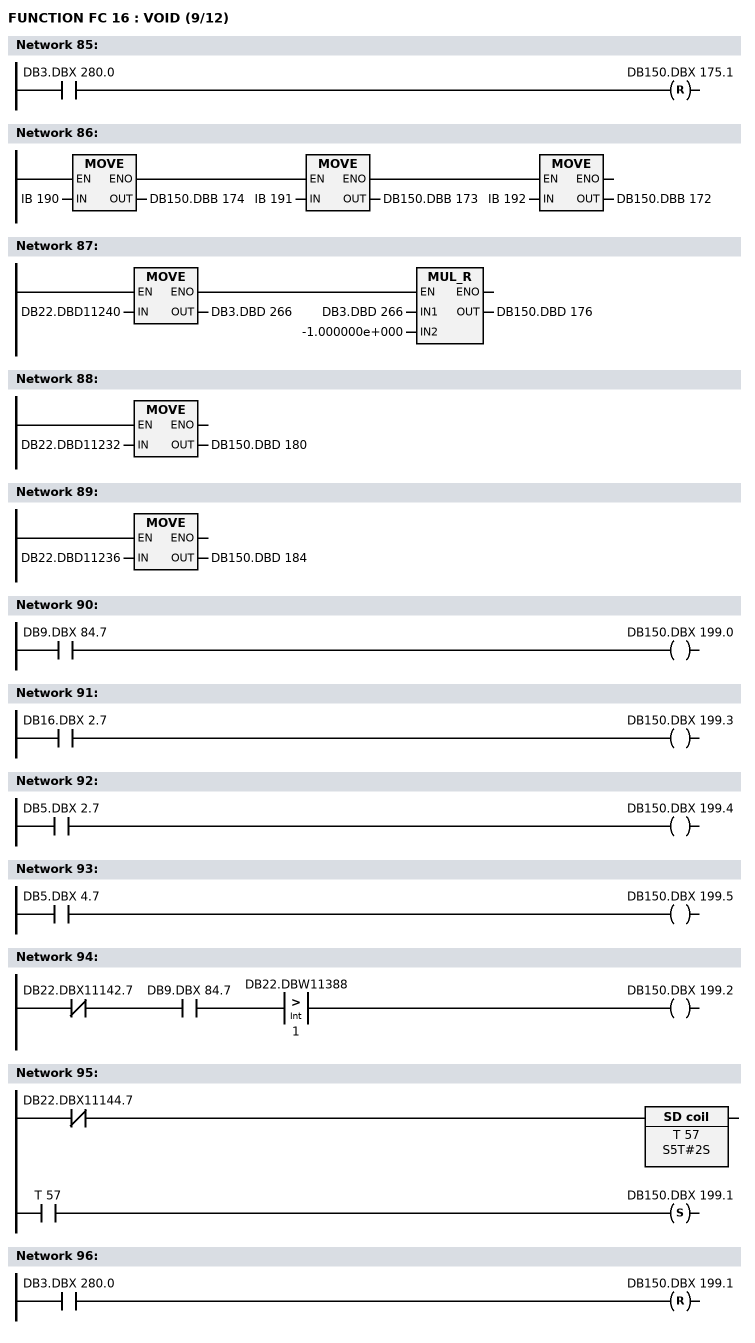

      A     DB3.DBX  280.0;
      R     DB150.DBX  175.1;
NETWORK
TITLE =

      A(    ;
      A(    ;
      L     IB   190;
      T     DB150.DBB  174;
      SET   ;
      SAVE  ;
      CLR   ;
      A     BR;
      )     ;
      JNB   M014;
      L     IB   191;
      T     DB150.DBB  173;
      SET   ;
      SAVE  ;
      CLR   ;
M014: A     BR;
      )     ;
      JNB   M015;
      L     IB   192;
      T     DB150.DBB  172;
M015: NOP   0;
NETWORK
TITLE =

      A(    ;
      L     DB22.DBD11240;
      T     DB3.DBD  266;
      SET   ;
      SAVE  ;
      CLR   ;
      A     BR;
      )     ;
      JNB   M016;
      L     DB3.DBD  266;
      L     -1.000000e+000;
      *R    ;
      T     DB150.DBD  176;
M016: NOP   0;
NETWORK
TITLE =

      L     DB22.DBD11232;
      T     DB150.DBD  180;
      NOP   0;
NETWORK
TITLE =

      L     DB22.DBD11236;
      T     DB150.DBD  184;
      NOP   0;
NETWORK
TITLE =

      A     DB9.DBX   84.7;
      =     DB150.DBX  199.0;
NETWORK
TITLE =

      A     DB16.DBX    2.7;
      =     DB150.DBX  199.3;
NETWORK
TITLE =

      A     DB5.DBX    2.7;
      =     DB150.DBX  199.4;
NETWORK
TITLE =

      A     DB5.DBX    4.7;
      =     DB150.DBX  199.5;
NETWORK
TITLE =

      AN    DB22.DBX11142.7;
      A     DB9.DBX   84.7;
      A(    ;
      L     DB22.DBW11388;
      L     1;
      >I    ;
      )     ;
      =     DB150.DBX  199.2;
NETWORK
TITLE =

      AN    DB22.DBX11144.7;
      L     S5T#2S;
      SD    T     57;
      NOP   0;
      NOP   0;
      NOP   0;
      A     T     57;
      S     DB150.DBX  199.1;
NETWORK
TITLE =

      A     DB3.DBX  280.0;
      R     DB150.DBX  199.1;
NETWORK
TITLE =
